	ELSIF TRUE 	
	AND fbPis.m_CheckByRecipe(stPis:=stPis_Tank_Water, 			req:=E_Piston_Recipe_State.Release)
	AND fbPis.m_CheckByRecipe(stPis:=stPis_Tank_R_Water, 		req:=E_Piston_Recipe_State.Release)
	AND fbPis.m_CheckByRecipe(stPis:=stPis_Tank_Detergent, 		req:=E_Piston_Recipe_State.Release)
	AND fbPis.m_CheckByRecipe(stPis:=stPis_Tank_DisInfection, 	req:=E_Piston_Recipe_State.Act)
	AND fbPis.m_CheckByRecipe(stPis:=stPis_Drain, 				req:=E_Piston_Recipe_State.Act)
	THEN;
		eStatus:=E_CIP_Source.eT91_Sanitation;
	ELSE;
		eStatus:=E_CIP_Source.eNone;
	END_IF
ELSE;
	eStatus:=E_CIP_Source.eNone;
END_IF
END_ACTION

METHOD m_CheckStatus : BOOL
VAR_INPUT
	eReqStatus		: E_CIP_Source;
END_VAR
IF eStatus=eReqStatus 
AND eProcess=E_CIP_Source.eNone
AND eReq=E_CIP_Source.eNone
AND bReady
AND bDone
AND NOT bRun
THEN;
	m_CheckStatus:=TRUE;
END_IF
END_METHOD

METHOD m_IsFree : BOOL
// In Ready with no request: a command given now will not be lost
IF eProcess=E_CIP_Source.eNone
AND eReq=E_CIP_Source.eNone
AND bReady
AND NOT bRun
THEN;
	m_IsFree:=TRUE;
END_IF
END_METHOD

METHOD m_Request_Reset : BOOL
VAR_IN_OUT
	memo: R_TRIG;
END_VAR
memo(CLK:=eReq=0);
IF TRUE 
AND memo.Q
THEN;
	SFCReset:=TRUE;
END_IF
END_METHOD

METHOD m_Run : BOOL
VAR_INPUT
	eReqProc			: E_CIP_Source;
END_VAR
IF eProcess=E_CIP_Source.eNone THEN;
	eProcess:=eReq:=eReqProc;
	bDone:=FALSE;
	m_Run:=TRUE;
END_IF
END_METHOD

METHOD m_Set_SFCFlags_Reference : BOOL
//Set reference to SFC flags

refSFC.SFCInit REF= SFCInit;
refSFC.SFCReset REF= SFCReset;
refSFC.SFCError REF= SFCError;
refSFC.SFCEnableLimit REF= SFCEnableLimit;
refSFC.SFCErrorStep REF= SFCErrorStep;
refSFC.SFCErrorPOU REF= SFCErrorPOU;
refSFC.SFCQuitError REF= SFCQuitError;
refSFC.SFCPause REF= SFCPause;
refSFC.SFCTrans REF= SFCTrans;
refSFC.SFCCurrentStep REF= SFCCurrentStep;
refSFC.SFCTip REF= SFCTip;
refSFC.SFCTipMode REF= SFCTipMode;

// Cycle handle for SFC
m_SFC_Handle();
END_METHOD

END_FUNCTION_BLOCK

// ---- 00 Library/03 SFC/FB_SFC_Cycle.TcPOU
FUNCTION_BLOCK FB_SFC_Cycle
VAR_INPUT

END_VAR
VAR_OUTPUT
END_VAR
VAR
	refSFC: ST_SFC;

	bInit: BOOL;
	bResetCycle: BOOL;
	bResume: BOOL;
	bRun: BOOL;	
	bReady: BOOL;
	bDone: BOOL;
	bToBe_Done: BOOL;
	
	bStepMode: BOOL;
	bNextStep: BOOL;



	bStepDone: BOOL;
	ton_StepTime: TON;
	
	StageDelayByRecipe: TIME;
	
	//fbPis_Meth: FB_Piston;

	rtDone	: R_TRIG;
	rtRun	: R_TRIG;
	sLastStepBefore_Error	: STRING;
	sError_Message			: STRING;
	
	ErrorSFC: BOOL;

	tonResetCycle: TON;
	
	stMode_zone	: REFERENCE TO ST_Mode;
	stOper_zone	: REFERENCE TO ST_OperationButtons;
	ftStateSafe : F_TRIG;
	
END_VAR

METHOD m_Reset_LastStepBeforeError : BOOL
VAR_INPUT
END_VAR
sLastStepBefore_Error:='';
END_METHOD

METHOD m_Set_LastStepBeforeError : BOOL
VAR_INPUT
END_VAR
sLastStepBefore_Error:=refSFC.SFCCurrentStep;
END_METHOD

METHOD m_Set_Mode_Reference : BOOL
VAR_INPUT
	inMoedeZone: E_ModeZone;
END_VAR
stMode_zone REF=(stMode[inMoedeZone]);
stOper_zone REF=(stOper[inMoedeZone]);
END_METHOD

METHOD m_SFC_Handle : BOOL
VAR_INPUT
END_VAR

VAR
	
END_VAR
IF NOT __ISVALIDREF(refSFC.SFCInit) 
OR NOT  __ISVALIDREF(refSFC.SFCReset) 
OR NOT  __ISVALIDREF(refSFC.SFCError) 
OR NOT  __ISVALIDREF(refSFC.SFCEnableLimit) 
OR NOT  __ISVALIDREF(refSFC.SFCErrorStep) 
OR NOT  __ISVALIDREF(refSFC.SFCErrorPOU) 
OR NOT  __ISVALIDREF(refSFC.SFCQuitError) 
OR NOT  __ISVALIDREF(refSFC.SFCPause) 
OR NOT  __ISVALIDREF(refSFC.SFCTrans) 
OR NOT  __ISVALIDREF(refSFC.SFCCurrentStep) 
OR NOT  __ISVALIDREF(refSFC.SFCTip) 
OR NOT  __ISVALIDREF(refSFC.SFCTipMode) 
THEN;
	RETURN;
END_IF

refSFC.SFCEnableLimit:=TRUE;
IF refSFC.SFCTrans THEN;
	bStepDone:=FALSE;
	ton_StepTime(IN:=FALSE);
ELSE;
	ton_StepTime(IN:=TRUE); //depend on step condition
END_IF

IF bInit THEN;
	refSFC.SFCInit:=TRUE;
ELSE;
	refSFC.SFCInit:=FALSE;
END_IF

IF refSFC.SFCError THEN;
	refSFC.SFCPause:=TRUE;
	ErrorSFC:=TRUE;
	m_Set_LastStepBeforeError();
END_IF

IF refSFC.SFCQuitError THEN;
	refSFC.SFCPause:=FALSE;
	ErrorSFC:=FALSE;
	refSFC.SFCQuitError:=FALSE;
	m_Reset_LastStepBeforeError();
	sError_Message:='';
END_IF

IF refSFC.SFCCurrentStep='Ready' THEN;
	bReady:=TRUE;
ELSE;
	bReady:=FALSE;
END_IF

rtDone(CLK:=refSFC.SFCCurrentStep='Done');
IF rtDone.Q THEN;
	bDone:=TRUE;
END_IF
rtRun(CLK:=bRun);
IF rtRun.Q THEN;
	bDone:=FALSE;
END_IF

IF bResume THEN;
	ErrorSFC:=FALSE;
	refSFC.SFCError:=FALSE;
	refSFC.SFCPause:=FALSE;
	m_Reset_LastStepBeforeError();
	bResume:=FALSE;
END_IF


tonResetCycle(PT:=T#0.5S,IN:=bResetCycle);
IF bResetCycle THEN;
	refSFC.SFCReset:=TRUE;
	//tonResetCycle.IN:=TRUE;
END_IF
IF tonResetCycle.Q THEN;
	bResetCycle:=FALSE;
	refSFC.SFCReset:=FALSE;
END_IF

StepByStep();

IF NOT __ISVALIDREF(stMode_zone)
OR NOT __ISVALIDREF(stOper_zone)
THEN;
	RETURN;
ELSE;
	//IF prg_Safety.ftStateSafe.Q THEN;
	ftStateSafe(CLK:=stMode_zone.bStateSafe_mode);
	IF ftStateSafe.Q THEN;
		//bResetCycle:=TRUE;
	END_IF	
END_IF



(*
rtDone(CLK:=bDone);
IF rtDone.Q THEN
	bToBe_Done:=FALSE;
END_IF
*)
END_METHOD

METHOD mInit : BOOL
VAR_INPUT
END_VAR
bInit:=TRUE;
bToBe_Done:=FALSE;
END_METHOD

METHOD mResetCycle : BOOL
VAR_INPUT
END_VAR
bResetCycle:=TRUE;
bRun:=FALSE;
refSFC.SFCReset:=TRUE;
END_METHOD

METHOD mRun : BOOL
VAR_INPUT
	
END_VAR
bRun:=TRUE;
bDone:=FALSE;

IF rtDone.Q THEN;
	mRun:=TRUE;	
END_IF
END_METHOD

METHOD mToBe_Done : BOOL
VAR_INPUT
END_VAR
bToBe_Done:=TRUE;
bDone:=FALSE;
END_METHOD

METHOD StepByStep : BOOL
VAR_INPUT
END_VAR


IF bStepMode THEN;
	IF refSFC.SFCTrans THEN;
		refSFC.SFCTipMode:=TRUE;
		bNextStep:=FALSE;
	END_IF
	IF bNextStep THEN;
		refSFC.SFCTipMode:=FALSE;
	END_IF
ELSE;
	refSFC.SFCTipMode:=FALSE;
END_IF
END_METHOD

END_FUNCTION_BLOCK

// ---- 03 Project/23 CIP/FB_CIP_Return.TcPOU
FUNCTION_BLOCK FB_CIP_Return EXTENDS FB_SFC_Cycle IMPLEMENTS ITF_FB_SFC_Cycle
VAR_INPUT
	//eElementID			: E_Element_List;
	
	valTank_Water			: E_Pis_Name;
	valTank_Water_1			: E_Pis_Name;
	valTank_R_Water			: E_Pis_Name;
	valTank_R_Water_1		: E_Pis_Name;
	valTank_Detergent		: E_Pis_Name;
	valTank_Detergent_1		: E_Pis_Name;
	valTank_DisInfection	: E_Pis_Name;
	valTank_DisInfection_1	: E_Pis_Name;
	valDrain				: E_Pis_Name;
	
END_VAR
VAR_OUTPUT
END_VAR
VAR
	//refElement		: REFERENCE TO FB_Element;
	//refState_Long		: REFERENCE TO E_Element_State_Long;
	eReq				: E_CIP_Return;
	eProcess			: E_CIP_Return;
	eStatus				: E_CIP_Return;
	
	fbPis						: FB_Piston;
	stPis_Tank_Water			: REFERENCE TO ST_Piston;
	stPis_Tank_Water_1			: REFERENCE TO ST_Piston;
	stPis_Tank_R_Water			: REFERENCE TO ST_Piston;
	stPis_Tank_R_Water_1		: REFERENCE TO ST_Piston;
	stPis_Tank_Detergent		: REFERENCE TO ST_Piston;
	stPis_Tank_Detergent_1		: REFERENCE TO ST_Piston;
	stPis_Tank_DisInfection		: REFERENCE TO ST_Piston;
	stPis_Tank_DisInfection_1	: REFERENCE TO ST_Piston;
	stPis_Drain					: REFERENCE TO ST_Piston;
	rt_Req_Reset: R_TRIG;
END_VAR
VAR_IN_OUT


END_VAR

act_GetReference();

act_Oper();
IF NOT Init.x THEN;
	act_Status();
END_IF

m_Request_Reset(memo:=rt_Req_Reset);//

ACTION _aDetergent_active:
bStepDone:=FALSE;
IF TRUE 
AND eStatus=E_CIP_Return.eT92_Detergent
THEN;
	bStepDone:=TRUE;
END_IF
END_ACTION

ACTION _aDetergent_entry:
fbPis.m_SetByRecipe(stPis:=stPis_Tank_Water, 			req:=E_Piston_Recipe_State.Release);
fbPis.m_SetByRecipe(stPis:=stPis_Tank_Water_1, 			req:=E_Piston_Recipe_State.Release);
fbPis.m_SetByRecipe(stPis:=stPis_Tank_R_Water, 			req:=E_Piston_Recipe_State.Release);
fbPis.m_SetByRecipe(stPis:=stPis_Tank_R_Water_1, 		req:=E_Piston_Recipe_State.Release);
fbPis.m_SetByRecipe(stPis:=stPis_Tank_Detergent, 		req:=E_Piston_Recipe_State.Act);
fbPis.m_SetByRecipe(stPis:=stPis_Tank_Detergent_1, 		req:=E_Piston_Recipe_State.Act);
fbPis.m_SetByRecipe(stPis:=stPis_Tank_DisInfection_1, 	req:=E_Piston_Recipe_State.Release);
fbPis.m_SetByRecipe(stPis:=stPis_Tank_DisInfection, 	req:=E_Piston_Recipe_State.Release);
fbPis.m_SetByRecipe(stPis:=stPis_Drain, 				req:=E_Piston_Recipe_State.Release);
END_ACTION

ACTION _aDone_entry:
eProcess:=E_CIP_Return.eNone; 
eReq:=E_CIP_Return.eNone;
bRun:=FALSE;
bDone:=TRUE;
END_ACTION

ACTION _aDrain_active:
bStepDone:=FALSE;
IF TRUE 
AND eStatus=E_CIP_Return.eDrain
THEN;
	bStepDone:=TRUE;
END_IF
END_ACTION

ACTION _aDrain_entry:
fbPis.m_SetByRecipe(stPis:=stPis_Tank_Water, 			req:=E_Piston_Recipe_State.Release);
fbPis.m_SetByRecipe(stPis:=stPis_Tank_Water_1, 			req:=E_Piston_Recipe_State.Release);
fbPis.m_SetByRecipe(stPis:=stPis_Tank_R_Water, 			req:=E_Piston_Recipe_State.Release);
fbPis.m_SetByRecipe(stPis:=stPis_Tank_R_Water_1, 		req:=E_Piston_Recipe_State.Release);
fbPis.m_SetByRecipe(stPis:=stPis_Tank_Detergent, 		req:=E_Piston_Recipe_State.Release);
fbPis.m_SetByRecipe(stPis:=stPis_Tank_Detergent_1, 		req:=E_Piston_Recipe_State.Release);
fbPis.m_SetByRecipe(stPis:=stPis_Tank_DisInfection, 	req:=E_Piston_Recipe_State.Release);
fbPis.m_SetByRecipe(stPis:=stPis_Tank_DisInfection_1, 	req:=E_Piston_Recipe_State.Release);
fbPis.m_SetByRecipe(stPis:=stPis_Drain, 				req:=E_Piston_Recipe_State.Release);
END_ACTION

ACTION _aInit_active:
SFCReset:=FALSE;
END_ACTION

ACTION _aInit_exit:
eProcess:=E_CIP_Return.eNone;
eReq:=E_CIP_Return.eNone;
END_ACTION

ACTION _aR_Water_active:
bStepDone:=FALSE;
IF TRUE 
AND eStatus=E_CIP_Return.eT93_R_Water
THEN;
	bStepDone:=TRUE;
END_IF
END_ACTION

ACTION _aR_Water_entry:
fbPis.m_SetByRecipe(stPis:=stPis_Tank_Water, 			req:=E_Piston_Recipe_State.Release);
fbPis.m_SetByRecipe(stPis:=stPis_Tank_Water_1, 			req:=E_Piston_Recipe_State.Release);
fbPis.m_SetByRecipe(stPis:=stPis_Tank_R_Water, 			req:=E_Piston_Recipe_State.Act);
fbPis.m_SetByRecipe(stPis:=stPis_Tank_R_Water_1, 		req:=E_Piston_Recipe_State.Act);
fbPis.m_SetByRecipe(stPis:=stPis_Tank_Detergent, 		req:=E_Piston_Recipe_State.Release);
fbPis.m_SetByRecipe(stPis:=stPis_Tank_Detergent_1, 		req:=E_Piston_Recipe_State.Release);
fbPis.m_SetByRecipe(stPis:=stPis_Tank_DisInfection, 	req:=E_Piston_Recipe_State.Release);
fbPis.m_SetByRecipe(stPis:=stPis_Tank_DisInfection_1, 	req:=E_Piston_Recipe_State.Release);
fbPis.m_SetByRecipe(stPis:=stPis_Drain, 				req:=E_Piston_Recipe_State.Release);
END_ACTION

ACTION _aReady_active:


CASE eReq OF
	E_CIP_Return.eDrain:;
			IF TRUE THEN;
				eProcess:=E_CIP_Return.eDrain;
			END_IF

	E_CIP_Return.eT91_Sanitation:;
			IF TRUE THEN;
				eProcess:=E_CIP_Return.eT91_Sanitation;
			END_IF	
			
	E_CIP_Return.eT92_Detergent:;
			IF TRUE THEN;
				eProcess:=E_CIP_Return.eT92_Detergent;
			END_IF	

	E_CIP_Return.eT93_R_Water:;
			IF TRUE THEN;
				eProcess:=E_CIP_Return.eT93_R_Water;
			END_IF	
			
	E_CIP_Return.eT94_Water:;
			IF TRUE THEN;
				eProcess:=E_CIP_Return.eT94_Water;
			END_IF	

END_CASE
END_ACTION

ACTION _aReady_entry:

END_ACTION

ACTION _aReady_exit:
bRun:=TRUE;
bDone:=FALSE;
END_ACTION

ACTION _aSanitation_active:
bStepDone:=FALSE;
IF TRUE 
AND eStatus=E_CIP_Return.eT91_Sanitation
THEN;
	bStepDone:=TRUE;
END_IF
END_ACTION

ACTION _aSanitation_entry:
fbPis.m_SetByRecipe(stPis:=stPis_Tank_Water, 			req:=E_Piston_Recipe_State.Release);
fbPis.m_SetByRecipe(stPis:=stPis_Tank_Water_1, 			req:=E_Piston_Recipe_State.Release);
fbPis.m_SetByRecipe(stPis:=stPis_Tank_R_Water, 			req:=E_Piston_Recipe_State.Release);
fbPis.m_SetByRecipe(stPis:=stPis_Tank_R_Water_1, 		req:=E_Piston_Recipe_State.Release);
fbPis.m_SetByRecipe(stPis:=stPis_Tank_Detergent, 		req:=E_Piston_Recipe_State.Release);
fbPis.m_SetByRecipe(stPis:=stPis_Tank_Detergent_1, 		req:=E_Piston_Recipe_State.Release);
fbPis.m_SetByRecipe(stPis:=stPis_Tank_DisInfection, 	req:=E_Piston_Recipe_State.Act);
fbPis.m_SetByRecipe(stPis:=stPis_Tank_DisInfection_1, 	req:=E_Piston_Recipe_State.Act);
fbPis.m_SetByRecipe(stPis:=stPis_Drain, 				req:=E_Piston_Recipe_State.Release);
END_ACTION

ACTION _aWater_active:
bStepDone:=FALSE;
IF TRUE 
AND eStatus=E_CIP_Return.eT94_Water
THEN;
	bStepDone:=TRUE;
END_IF
END_ACTION

ACTION _aWater_entry:
fbPis.m_SetByRecipe(stPis:=stPis_Tank_Water, 			req:=E_Piston_Recipe_State.Act);
fbPis.m_SetByRecipe(stPis:=stPis_Tank_Water_1, 			req:=E_Piston_Recipe_State.Act);
fbPis.m_SetByRecipe(stPis:=stPis_Tank_R_Water, 			req:=E_Piston_Recipe_State.Release);
fbPis.m_SetByRecipe(stPis:=stPis_Tank_R_Water_1, 		req:=E_Piston_Recipe_State.Release);
fbPis.m_SetByRecipe(stPis:=stPis_Tank_Detergent, 		req:=E_Piston_Recipe_State.Release);
fbPis.m_SetByRecipe(stPis:=stPis_Tank_Detergent_1, 		req:=E_Piston_Recipe_State.Release);
fbPis.m_SetByRecipe(stPis:=stPis_Tank_DisInfection, 	req:=E_Piston_Recipe_State.Release);
fbPis.m_SetByRecipe(stPis:=stPis_Tank_DisInfection_1, 	req:=E_Piston_Recipe_State.Release);
fbPis.m_SetByRecipe(stPis:=stPis_Drain, 				req:=E_Piston_Recipe_State.Act);
END_ACTION

ACTION act_GetReference:
m_Set_SFCFlags_Reference();
//refElement REF= fbElement[eElementID];
//refState_Long REF= fbElement[eElementID].eState_Long;
	
stPis_Tank_Water				REF= g_Piston.stPis[valTank_Water];
stPis_Tank_Water_1				REF= g_Piston.stPis[valTank_Water_1];
stPis_Tank_R_Water				REF= g_Piston.stPis[valTank_R_Water];
stPis_Tank_R_Water_1			REF= g_Piston.stPis[valTank_R_Water_1];
stPis_Tank_Detergent			REF= g_Piston.stPis[valTank_Detergent];
stPis_Tank_Detergent_1			REF= g_Piston.stPis[valTank_Detergent_1];
stPis_Tank_DisInfection			REF= g_Piston.stPis[valTank_DisInfection];
stPis_Tank_DisInfection_1		REF= g_Piston.stPis[valTank_DisInfection_1];
stPis_Drain						REF= g_Piston.stPis[valDrain];
END_ACTION

ACTION act_Oper:
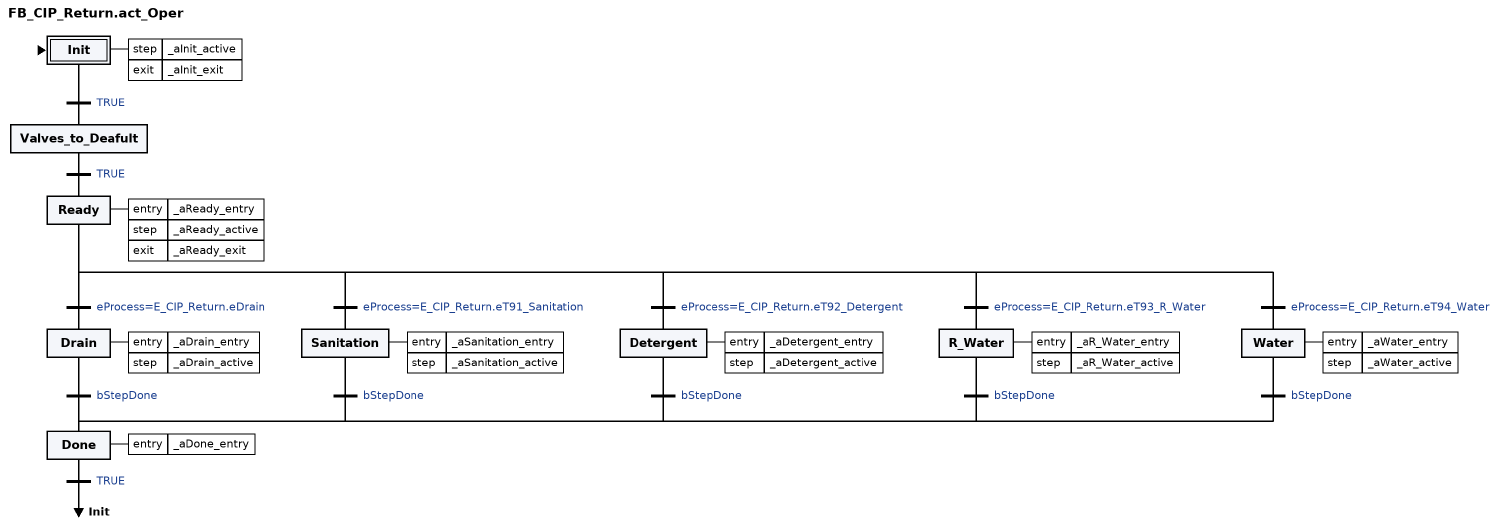
INITIAL_STEP Init:  // min time T#0.5s
    _aInit_active(N);  // step action
    _aInit_exit(P0);  // exit action
END_STEP
TRANSITION FROM Init TO Valves_to_Deafult
    := TRUE;
END_TRANSITION
STEP Valves_to_Deafult:
END_STEP
TRANSITION FROM Valves_to_Deafult TO Ready
    := TRUE;
END_TRANSITION
STEP Ready:
    _aReady_entry(P1);  // entry action
    _aReady_active(N);  // step action
    _aReady_exit(P0);  // exit action
END_STEP
TRANSITION FROM Ready TO Drain
    := eProcess=E_CIP_Return.eDrain;
END_TRANSITION
STEP Drain:
    _aDrain_entry(P1);  // entry action
    _aDrain_active(N);  // step action
END_STEP
TRANSITION FROM Drain TO Done
    := bStepDone;
END_TRANSITION
TRANSITION FROM Ready TO Sanitation
    := eProcess=E_CIP_Return.eT91_Sanitation;
END_TRANSITION
STEP Sanitation:
    _aSanitation_entry(P1);  // entry action
    _aSanitation_active(N);  // step action
END_STEP
TRANSITION FROM Sanitation TO Done
    := bStepDone;
END_TRANSITION
TRANSITION FROM Ready TO Detergent
    := eProcess=E_CIP_Return.eT92_Detergent;
END_TRANSITION
STEP Detergent:
    _aDetergent_entry(P1);  // entry action
    _aDetergent_active(N);  // step action
END_STEP
TRANSITION FROM Detergent TO Done
    := bStepDone;
END_TRANSITION
TRANSITION FROM Ready TO R_Water
    := eProcess=E_CIP_Return.eT93_R_Water;
END_TRANSITION
STEP R_Water:
    _aR_Water_entry(P1);  // entry action
    _aR_Water_active(N);  // step action
END_STEP
TRANSITION FROM R_Water TO Done
    := bStepDone;
END_TRANSITION
TRANSITION FROM Ready TO Water
    := eProcess=E_CIP_Return.eT94_Water;
END_TRANSITION
STEP Water:
    _aWater_entry(P1);  // entry action
    _aWater_active(N);  // step action
END_STEP
TRANSITION FROM Water TO Done
    := bStepDone;
END_TRANSITION
STEP Done:  // min time T#0.2s
    _aDone_entry(P1);  // entry action
END_STEP
TRANSITION FROM Done TO Init
    := TRUE;
END_TRANSITION
// branch label Branch1_act_Oper
END_ACTION

ACTION act_Status:
IF bReady AND bDone OR TRUE THEN;
	IF TRUE 
	AND fbPis.m_CheckByRecipe(stPis:=stPis_Tank_Water, 			req:=E_Piston_Recipe_State.Release)
	AND fbPis.m_CheckByRecipe(stPis:=stPis_Tank_R_Water, 		req:=E_Piston_Recipe_State.Release)
	AND fbPis.m_CheckByRecipe(stPis:=stPis_Tank_Detergent, 		req:=E_Piston_Recipe_State.Release)
	AND fbPis.m_CheckByRecipe(stPis:=stPis_Tank_DisInfection, 	req:=E_Piston_Recipe_State.Release)
	AND fbPis.m_CheckByRecipe(stPis:=stPis_Drain, 				req:=E_Piston_Recipe_State.Release)
	AND fbPis.m_CheckByRecipe(stPis:=stPis_Tank_Water_1, 		req:=E_Piston_Recipe_State.Release)
	AND fbPis.m_CheckByRecipe(stPis:=stPis_Tank_R_Water_1, 		req:=E_Piston_Recipe_State.Release)
	AND fbPis.m_CheckByRecipe(stPis:=stPis_Tank_Detergent_1, 	req:=E_Piston_Recipe_State.Release)
	AND fbPis.m_CheckByRecipe(stPis:=stPis_Tank_DisInfection_1, req:=E_Piston_Recipe_State.Release)
	THEN;
		eStatus:=E_CIP_Return.eDrain;
	
	ELSIF TRUE 
	AND fbPis.m_CheckByRecipe(stPis:=stPis_Tank_Water, 			req:=E_Piston_Recipe_State.Act)
	AND fbPis.m_CheckByRecipe(stPis:=stPis_Tank_R_Water, 		req:=E_Piston_Recipe_State.Release)
	AND fbPis.m_CheckByRecipe(stPis:=stPis_Tank_Detergent, 		req:=E_Piston_Recipe_State.Release)
	AND fbPis.m_CheckByRecipe(stPis:=stPis_Tank_DisInfection, 	req:=E_Piston_Recipe_State.Release)
	AND fbPis.m_CheckByRecipe(stPis:=stPis_Drain, 				req:=E_Piston_Recipe_State.Act)
	AND fbPis.m_CheckByRecipe(stPis:=stPis_Tank_Water_1, 		req:=E_Piston_Recipe_State.Act)
	AND fbPis.m_CheckByRecipe(stPis:=stPis_Tank_R_Water_1, 		req:=E_Piston_Recipe_State.Release)
	AND fbPis.m_CheckByRecipe(stPis:=stPis_Tank_Detergent_1, 	req:=E_Piston_Recipe_State.Release)
	AND fbPis.m_CheckByRecipe(stPis:=stPis_Tank_DisInfection_1, req:=E_Piston_Recipe_State.Release)
	THEN;
		eStatus:=E_CIP_Return.eT94_Water;
		
	ELSIF TRUE 
	AND fbPis.m_CheckByRecipe(stPis:=stPis_Tank_Water, 			req:=E_Piston_Recipe_State.Release)
	AND fbPis.m_CheckByRecipe(stPis:=stPis_Tank_R_Water, 		req:=E_Piston_Recipe_State.Act)
	AND fbPis.m_CheckByRecipe(stPis:=stPis_Tank_Detergent, 		req:=E_Piston_Recipe_State.Release)
	AND fbPis.m_CheckByRecipe(stPis:=stPis_Tank_DisInfection, 	req:=E_Piston_Recipe_State.Release)
	AND fbPis.m_CheckByRecipe(stPis:=stPis_Drain, 				req:=E_Piston_Recipe_State.Release)
	AND fbPis.m_CheckByRecipe(stPis:=stPis_Tank_Water_1, 			req:=E_Piston_Recipe_State.Release)
	AND fbPis.m_CheckByRecipe(stPis:=stPis_Tank_R_Water_1, 			req:=E_Piston_Recipe_State.Act)
	AND fbPis.m_CheckByRecipe(stPis:=stPis_Tank_Detergent_1, 		req:=E_Piston_Recipe_State.Release)
	AND fbPis.m_CheckByRecipe(stPis:=stPis_Tank_DisInfection_1, 	req:=E_Piston_Recipe_State.Release)
	THEN;
		eStatus:=E_CIP_Return.eT93_R_Water;
		
	ELSIF TRUE 	
	AND fbPis.m_CheckByRecipe(stPis:=stPis_Tank_Water, 			req:=E_Piston_Recipe_State.Release)
	AND fbPis.m_CheckByRecipe(stPis:=stPis_Tank_R_Water, 		req:=E_Piston_Recipe_State.Release)
	AND fbPis.m_CheckByRecipe(stPis:=stPis_Tank_Detergent, 		req:=E_Piston_Recipe_State.Act)
	AND fbPis.m_CheckByRecipe(stPis:=stPis_Tank_DisInfection, 	req:=E_Piston_Recipe_State.Release)
	AND fbPis.m_CheckByRecipe(stPis:=stPis_Drain, 				req:=E_Piston_Recipe_State.Release)
	AND fbPis.m_CheckByRecipe(stPis:=stPis_Tank_Water_1, 			req:=E_Piston_Recipe_State.Release)
	AND fbPis.m_CheckByRecipe(stPis:=stPis_Tank_R_Water_1, 			req:=E_Piston_Recipe_State.Release)
	AND fbPis.m_CheckByRecipe(stPis:=stPis_Tank_Detergent_1, 		req:=E_Piston_Recipe_State.Act)
	AND fbPis.m_CheckByRecipe(stPis:=stPis_Tank_DisInfection_1, 	req:=E_Piston_Recipe_State.Release)
	THEN;
		eStatus:=E_CIP_Return.eT92_Detergent;
		
	ELSIF TRUE 	
	AND fbPis.m_CheckByRecipe(stPis:=stPis_Tank_Water, 			req:=E_Piston_Recipe_State.Release)
	AND fbPis.m_CheckByRecipe(stPis:=stPis_Tank_R_Water, 		req:=E_Piston_Recipe_State.Release)
	AND fbPis.m_CheckByRecipe(stPis:=stPis_Tank_Detergent, 		req:=E_Piston_Recipe_State.Release)
	AND fbPis.m_CheckByRecipe(stPis:=stPis_Tank_DisInfection, 	req:=E_Piston_Recipe_State.Act)
	AND fbPis.m_CheckByRecipe(stPis:=stPis_Drain, 				req:=E_Piston_Recipe_State.Release)
	AND fbPis.m_CheckByRecipe(stPis:=stPis_Tank_Water_1, 			req:=E_Piston_Recipe_State.Release)
	AND fbPis.m_CheckByRecipe(stPis:=stPis_Tank_R_Water_1, 			req:=E_Piston_Recipe_State.Release)
	AND fbPis.m_CheckByRecipe(stPis:=stPis_Tank_Detergent_1, 		req:=E_Piston_Recipe_State.Release)
	AND fbPis.m_CheckByRecipe(stPis:=stPis_Tank_DisInfection_1, 	req:=E_Piston_Recipe_State.Act)
	THEN;
		eStatus:=E_CIP_Return.eT91_Sanitation;
	ELSE;
		eStatus:=E_CIP_Return.eNone;
	END_IF
ELSE;
	eStatus:=E_CIP_Return.eNone;
END_IF
END_ACTION

METHOD m_CheckStatus : BOOL
VAR_INPUT
	eReqStatus		: E_CIP_Return;
END_VAR
IF eStatus=eReqStatus 
AND eProcess=E_CIP_Return.eNone
AND eReq=E_CIP_Return.eNone
AND bReady
AND bDone
AND NOT bRun
THEN;
	m_CheckStatus:=TRUE;
END_IF
END_METHOD

METHOD m_IsFree : BOOL
// In Ready with no request: a command given now will not be lost
IF eProcess=E_CIP_Return.eNone
AND eReq=E_CIP_Return.eNone
AND bReady
AND NOT bRun
THEN;
	m_IsFree:=TRUE;
END_IF
END_METHOD

METHOD m_Request_Reset : BOOL
VAR_IN_OUT
	memo: R_TRIG;
END_VAR
memo(CLK:=eReq=0);
IF TRUE 
AND memo.Q
THEN;
	SFCReset:=TRUE;
END_IF
END_METHOD

METHOD m_Run : BOOL
VAR_INPUT
	eReqProc			: E_CIP_Return;
END_VAR
IF eProcess=E_CIP_Return.eNone THEN;
	eProcess:=eReq:=eReqProc;
	bDone:=FALSE;
	m_Run:=TRUE;
END_IF
END_METHOD

METHOD m_Set_SFCFlags_Reference : BOOL
//Set reference to SFC flags

refSFC.SFCInit REF= SFCInit;
refSFC.SFCReset REF= SFCReset;
refSFC.SFCError REF= SFCError;
refSFC.SFCEnableLimit REF= SFCEnableLimit;
refSFC.SFCErrorStep REF= SFCErrorStep;
refSFC.SFCErrorPOU REF= SFCErrorPOU;
refSFC.SFCQuitError REF= SFCQuitError;
refSFC.SFCPause REF= SFCPause;
refSFC.SFCTrans REF= SFCTrans;
refSFC.SFCCurrentStep REF= SFCCurrentStep;
refSFC.SFCTip REF= SFCTip;
refSFC.SFCTipMode REF= SFCTipMode;

// Cycle handle for SFC
m_SFC_Handle();
END_METHOD

END_FUNCTION_BLOCK

// ---- 03 Project/23 CIP/FB_CIP_Client.TcPOU
FUNCTION_BLOCK FB_CIP_Client EXTENDS FB_SFC_Cycle IMPLEMENTS ITF_FB_SFC_Cycle
VAR_INPUT
	//eElementID			: E_Element_List;
	
	valClient_Source		: E_Pis_Name;
	valClient_Return		: E_Pis_Name;
	valS_Marinade_Up		: E_Pis_Name;
	//valS_Marinade_Up_Drain	: E_Pis_Name;
	valS_Marinade_Low		: E_Pis_Name;
	valS_Color_Up			: E_Pis_Name;
	//valS_Color_Up_Drain		: E_Pis_Name;
	valS_Color_Low			: E_Pis_Name;
	//valTank_1				: E_Pis_Name;
	//valTank_2				: E_Pis_Name;
	//valTank_3				: E_Pis_Name;
	//valTank_4				: E_Pis_Name;
	//valS_Marinade_Low_Select	: E_Pis_Name;
	//valS_Color_Low_Select	: E_Pis_Name;
	valDrain				: E_Pis_Name;
	valLoop					: E_Pis_Name;//V1030
	valS_Future				: E_Pis_Name;
	
END_VAR
VAR_OUTPUT
END_VAR
VAR
	//refElement		: REFERENCE TO FB_Element;
	//refState_Long		: REFERENCE TO E_Element_State_Long;
	eReq				: E_CIP_Client_Selector;
	eProcess			: E_CIP_Client_Selector;
	eStatus				: E_CIP_Client_Selector;
	
	fbPis					: FB_Piston;
	stPis_Client_Source			: REFERENCE TO ST_Piston;
	stPis_Client_Return			: REFERENCE TO ST_Piston;
	stPis_S_Marinade_Up			: REFERENCE TO ST_Piston;
	//stPis_S_Marinade_Up_Drain	: REFERENCE TO ST_Piston;
	stPis_S_Marinade_Low		: REFERENCE TO ST_Piston;
	stPis_S_Color_Up			: REFERENCE TO ST_Piston;
	//stPis_S_Color_Up_Drain		: REFERENCE TO ST_Piston;
	stPis_S_Color_Low			: REFERENCE TO ST_Piston;
	//stPis_Tank_1				: REFERENCE TO ST_Piston;
	//stPis_Tank_2				: REFERENCE TO ST_Piston;
	//stPis_Tank_3				: REFERENCE TO ST_Piston;
	//stPis_Tank_4				: REFERENCE TO ST_Piston;
	//stPis_S_Marinade_Low_Select	: REFERENCE TO ST_Piston;
	//stPis_S_Color_Low_Select	: REFERENCE TO ST_Piston;
	stPis_Drain					: REFERENCE TO ST_Piston;	
	stPis_Loop					: REFERENCE TO ST_Piston;//V1030
	stPis_S_Future				: REFERENCE TO ST_Piston;

	tonDrainTime: TON;
	
	rt_Req_Reset: R_TRIG;

END_VAR
VAR_IN_OUT


END_VAR

act_GetReference();

act_Oper();
IF NOT Init.x THEN;
	act_Status();
END_IF

tonDrainTime(PT:=T#1M, IN:=eStatus=E_CIP_Client_Selector.eDrain);
IF tonDrainTime.Q 
AND eReq=E_CIP_Client_Selector.eNone
AND eProcess=E_CIP_Client_Selector.eNone
THEN;
	eReq:=E_CIP_Client_Selector.eClose;
END_IF

m_Request_Reset(memo:=rt_Req_Reset);//rt_Req_Reset: R_TRIG;

ACTION _aClose_active:
bStepDone:=FALSE;
IF TRUE 
AND eStatus=E_CIP_Client_Selector.eClose
THEN;
	bStepDone:=TRUE;
END_IF
END_ACTION

ACTION _aClose_entry:
fbPis.m_SetByRecipe(stPis:=stPis_Client_Source, 		req:=E_Piston_Recipe_State.Release);
fbPis.m_SetByRecipe(stPis:=stPis_Client_Return, 		req:=E_Piston_Recipe_State.Release);
fbPis.m_SetByRecipe(stPis:=stPis_S_Marinade_Up, 		req:=E_Piston_Recipe_State.Release);
fbPis.m_SetByRecipe(stPis:=stPis_S_Marinade_Low, 		req:=E_Piston_Recipe_State.Release);
fbPis.m_SetByRecipe(stPis:=stPis_S_Color_Up, 			req:=E_Piston_Recipe_State.Release);
fbPis.m_SetByRecipe(stPis:=stPis_S_Color_Low, 			req:=E_Piston_Recipe_State.Release);
fbPis.m_SetByRecipe(stPis:=stPis_Drain, 				req:=E_Piston_Recipe_State.Release);
fbPis.m_SetByRecipe(stPis:=stPis_Loop, 					req:=E_Piston_Recipe_State.Release);
fbPis.m_SetByRecipe(stPis:=stPis_S_Future, 				req:=E_Piston_Recipe_State.Release);
END_ACTION

ACTION _aColor_Low_active:
bStepDone:=FALSE;
IF TRUE 
AND eStatus=E_CIP_Client_Selector.eColor_Low
THEN;
	bStepDone:=TRUE;
END_IF
END_ACTION

ACTION _aColor_Low_entry:
fbPis.m_SetByRecipe(stPis:=stPis_Client_Source, 		req:=E_Piston_Recipe_State.Act);
fbPis.m_SetByRecipe(stPis:=stPis_Client_Return, 		req:=E_Piston_Recipe_State.Act);
fbPis.m_SetByRecipe(stPis:=stPis_S_Marinade_Up, 		req:=E_Piston_Recipe_State.Release);
fbPis.m_SetByRecipe(stPis:=stPis_S_Marinade_Low, 		req:=E_Piston_Recipe_State.Release);
fbPis.m_SetByRecipe(stPis:=stPis_S_Color_Up, 			req:=E_Piston_Recipe_State.Release);
fbPis.m_SetByRecipe(stPis:=stPis_S_Color_Low, 			req:=E_Piston_Recipe_State.Act);
fbPis.m_SetByRecipe(stPis:=stPis_Drain, 				req:=E_Piston_Recipe_State.Release);
fbPis.m_SetByRecipe(stPis:=stPis_Loop, 					req:=E_Piston_Recipe_State.Release);
fbPis.m_SetByRecipe(stPis:=stPis_S_Future, 				req:=E_Piston_Recipe_State.Release);
END_ACTION

ACTION _aColor_Up_active:
bStepDone:=FALSE;
IF TRUE 
AND eStatus=E_CIP_Client_Selector.eColor_Up
THEN;
	bStepDone:=TRUE;
END_IF
END_ACTION

ACTION _aColor_Up_entry:
fbPis.m_SetByRecipe(stPis:=stPis_Client_Source, 		req:=E_Piston_Recipe_State.Act);
fbPis.m_SetByRecipe(stPis:=stPis_Client_Return, 		req:=E_Piston_Recipe_State.Act);
fbPis.m_SetByRecipe(stPis:=stPis_S_Marinade_Up, 		req:=E_Piston_Recipe_State.Release);
fbPis.m_SetByRecipe(stPis:=stPis_S_Marinade_Low, 		req:=E_Piston_Recipe_State.Release);
fbPis.m_SetByRecipe(stPis:=stPis_S_Color_Up, 			req:=E_Piston_Recipe_State.Act);
fbPis.m_SetByRecipe(stPis:=stPis_S_Color_Low, 			req:=E_Piston_Recipe_State.Release);
fbPis.m_SetByRecipe(stPis:=stPis_Drain, 				req:=E_Piston_Recipe_State.Release);
fbPis.m_SetByRecipe(stPis:=stPis_Loop, 					req:=E_Piston_Recipe_State.Release);
fbPis.m_SetByRecipe(stPis:=stPis_S_Future, 				req:=E_Piston_Recipe_State.Release);
END_ACTION

ACTION _aDone_entry:
eProcess:=E_CIP_Usage.eNotInUse;
eReq:=E_CIP_Usage.eNotInUse;
bRun:=FALSE;
bDone:=TRUE;
END_ACTION

ACTION _aDrain_active:
bStepDone:=FALSE;
IF TRUE 
AND eStatus=E_CIP_Client_Selector.eDrain
THEN;
	bStepDone:=TRUE;
END_IF
END_ACTION

ACTION _aDrain_entry:
fbPis.m_SetByRecipe(stPis:=stPis_Client_Source, 		req:=E_Piston_Recipe_State.Release);
fbPis.m_SetByRecipe(stPis:=stPis_Client_Return, 		req:=E_Piston_Recipe_State.Release);
fbPis.m_SetByRecipe(stPis:=stPis_S_Marinade_Up, 		req:=E_Piston_Recipe_State.Release);
fbPis.m_SetByRecipe(stPis:=stPis_S_Marinade_Low, 		req:=E_Piston_Recipe_State.Release);
fbPis.m_SetByRecipe(stPis:=stPis_S_Color_Up, 			req:=E_Piston_Recipe_State.Release);
fbPis.m_SetByRecipe(stPis:=stPis_S_Color_Low, 			req:=E_Piston_Recipe_State.Release);
fbPis.m_SetByRecipe(stPis:=stPis_Drain, 				req:=E_Piston_Recipe_State.Act);
fbPis.m_SetByRecipe(stPis:=stPis_Loop, 					req:=E_Piston_Recipe_State.Release);
fbPis.m_SetByRecipe(stPis:=stPis_S_Future, 				req:=E_Piston_Recipe_State.Release);
END_ACTION

ACTION _aFuture_active:
bStepDone:=FALSE;
IF TRUE 
AND eStatus=E_CIP_Client_Selector.eFuture
THEN;
	bStepDone:=TRUE;
END_IF
END_ACTION

ACTION _aFuture_entry:
fbPis.m_SetByRecipe(stPis:=stPis_Client_Source, 		req:=E_Piston_Recipe_State.Act);
fbPis.m_SetByRecipe(stPis:=stPis_Client_Return, 		req:=E_Piston_Recipe_State.Act);
fbPis.m_SetByRecipe(stPis:=stPis_S_Marinade_Up, 		req:=E_Piston_Recipe_State.Release);
fbPis.m_SetByRecipe(stPis:=stPis_S_Marinade_Low, 		req:=E_Piston_Recipe_State.Release);
fbPis.m_SetByRecipe(stPis:=stPis_S_Color_Up, 			req:=E_Piston_Recipe_State.Release);
fbPis.m_SetByRecipe(stPis:=stPis_S_Color_Low, 			req:=E_Piston_Recipe_State.Release);
fbPis.m_SetByRecipe(stPis:=stPis_Drain, 				req:=E_Piston_Recipe_State.Release);
fbPis.m_SetByRecipe(stPis:=stPis_Loop, 					req:=E_Piston_Recipe_State.Release);
fbPis.m_SetByRecipe(stPis:=stPis_S_Future, 				req:=E_Piston_Recipe_State.Release);	//route to the plant: only source and return open
END_ACTION

ACTION _aInit_active:
SFCReset:=FALSE;
END_ACTION

ACTION _aInit_exit:
eProcess:=E_CIP_Usage.eNotInUse;
eReq:=E_CIP_Usage.eNotInUse;
END_ACTION

ACTION _aLoop_active:
bStepDone:=FALSE;
IF TRUE 
AND eStatus=E_CIP_Client_Selector.eLoop
THEN;
	bStepDone:=TRUE;
END_IF
END_ACTION

ACTION _aLoop_entry:
fbPis.m_SetByRecipe(stPis:=stPis_Client_Source, 		req:=E_Piston_Recipe_State.Act);
fbPis.m_SetByRecipe(stPis:=stPis_Client_Return, 		req:=E_Piston_Recipe_State.Act);
fbPis.m_SetByRecipe(stPis:=stPis_S_Marinade_Up, 		req:=E_Piston_Recipe_State.Release);
fbPis.m_SetByRecipe(stPis:=stPis_S_Marinade_Low, 		req:=E_Piston_Recipe_State.Release);
fbPis.m_SetByRecipe(stPis:=stPis_S_Color_Up, 			req:=E_Piston_Recipe_State.Release);
fbPis.m_SetByRecipe(stPis:=stPis_S_Color_Low, 			req:=E_Piston_Recipe_State.Release);
fbPis.m_SetByRecipe(stPis:=stPis_Drain, 				req:=E_Piston_Recipe_State.Act);
fbPis.m_SetByRecipe(stPis:=stPis_Loop, 					req:=E_Piston_Recipe_State.Act);
fbPis.m_SetByRecipe(stPis:=stPis_S_Future, 				req:=E_Piston_Recipe_State.Release);
END_ACTION

ACTION _aMarinade_Low_active:
bStepDone:=FALSE;
IF TRUE 
AND eStatus=E_CIP_Client_Selector.eMarinade_Low
THEN;
	bStepDone:=TRUE;
END_IF
END_ACTION

ACTION _aMarinade_Low_entry:
fbPis.m_SetByRecipe(stPis:=stPis_Client_Source, 		req:=E_Piston_Recipe_State.Act);
fbPis.m_SetByRecipe(stPis:=stPis_Client_Return, 		req:=E_Piston_Recipe_State.Act);
fbPis.m_SetByRecipe(stPis:=stPis_S_Marinade_Up, 		req:=E_Piston_Recipe_State.Release);
fbPis.m_SetByRecipe(stPis:=stPis_S_Marinade_Low, 		req:=E_Piston_Recipe_State.Act);
fbPis.m_SetByRecipe(stPis:=stPis_S_Color_Up, 			req:=E_Piston_Recipe_State.Release);
fbPis.m_SetByRecipe(stPis:=stPis_S_Color_Low, 			req:=E_Piston_Recipe_State.Release);
fbPis.m_SetByRecipe(stPis:=stPis_Drain, 				req:=E_Piston_Recipe_State.Release);
fbPis.m_SetByRecipe(stPis:=stPis_Loop, 					req:=E_Piston_Recipe_State.Release);
fbPis.m_SetByRecipe(stPis:=stPis_S_Future, 				req:=E_Piston_Recipe_State.Release);
END_ACTION

ACTION _aMarinade_Up_active:
bStepDone:=FALSE;
IF TRUE 
AND eStatus=E_CIP_Client_Selector.eMarinade_Up
THEN;
	bStepDone:=TRUE;
END_IF
END_ACTION

ACTION _aMarinade_Up_entry:
fbPis.m_SetByRecipe(stPis:=stPis_Client_Source, 		req:=E_Piston_Recipe_State.Act);
fbPis.m_SetByRecipe(stPis:=stPis_Client_Return, 		req:=E_Piston_Recipe_State.Act);
fbPis.m_SetByRecipe(stPis:=stPis_S_Marinade_Up, 		req:=E_Piston_Recipe_State.Act);
fbPis.m_SetByRecipe(stPis:=stPis_S_Marinade_Low, 		req:=E_Piston_Recipe_State.Release);
fbPis.m_SetByRecipe(stPis:=stPis_S_Color_Up, 			req:=E_Piston_Recipe_State.Release);
fbPis.m_SetByRecipe(stPis:=stPis_S_Color_Low, 			req:=E_Piston_Recipe_State.Release);
fbPis.m_SetByRecipe(stPis:=stPis_Drain, 				req:=E_Piston_Recipe_State.Release);
fbPis.m_SetByRecipe(stPis:=stPis_Loop, 					req:=E_Piston_Recipe_State.Release);
fbPis.m_SetByRecipe(stPis:=stPis_S_Future, 				req:=E_Piston_Recipe_State.Release);
END_ACTION

ACTION _aReady_active:


IF eReq<>E_CIP_Client_Selector.eNone THEN;
	IF eProcess=E_CIP_Client_Selector.eNone 
	THEN;
		eProcess:=eReq;
	ELSE;
		eReq:=E_CIP_Client_Selector.eNone;
	END_IF
END_IF

(*
CASE eReq OF
	E_CIP_Usage.eLine_Color:;
			IF TRUE THEN;
				eProcess:=E_CIP_Usage.eLine_Color;
			END_IF

	E_CIP_Usage.eLine_Marinada:;
			IF TRUE THEN;
				eProcess:=E_CIP_Usage.eLine_Marinada;
			END_IF	
			
	E_CIP_Usage.eLocal:;
			IF TRUE THEN;
				eProcess:=E_CIP_Usage.eLocal;
			END_IF	

	E_CIP_Usage.eNotInUse:;
			IF TRUE THEN;
				eProcess:=E_CIP_Usage.eNotInUse;
			END_IF	
			
	E_CIP_Usage.eTank_1:;
			IF TRUE THEN;
				eProcess:=E_CIP_Usage.eTank_1;
			END_IF	
	E_CIP_Usage.eTank_2:;
			IF TRUE THEN;
				eProcess:=E_CIP_Usage.eTank_2;
			END_IF	
	E_CIP_Usage.eTank_3:;
			IF TRUE THEN;
				eProcess:=E_CIP_Usage.eTank_3;
			END_IF	
	E_CIP_Usage.eTank_4:;
			IF TRUE THEN;
				eProcess:=E_CIP_Usage.eTank_4;
			END_IF	
	E_CIP_Usage.eTriBlender_Color:;
			IF TRUE THEN;
				eProcess:=E_CIP_Usage.eTriBlender_Color;
			END_IF	
	E_CIP_Usage.eTriBlender_Marinada:;
			IF TRUE THEN;
				eProcess:=E_CIP_Usage.eTriBlender_Marinada;
			END_IF	

END_CASE
*)
END_ACTION

ACTION _aReady_exit:
bRun:=TRUE;
bDone:=FALSE;
END_ACTION

ACTION act_GetReference:
m_Set_SFCFlags_Reference();
//refElement REF= fbElement[eElementID];
//refState_Long REF= fbElement[eElementID].eState_Long;

stPis_Client_Source			REF= g_Piston.stPis[valClient_Source];
stPis_Client_Return			REF= g_Piston.stPis[valClient_Return];
stPis_S_Marinade_Up			REF= g_Piston.stPis[valS_Marinade_Up];
//stPis_S_Marinade_Up_Drain	REF= g_Piston.stPis[valS_Marinade_Up_Drain];
stPis_S_Marinade_Low		REF= g_Piston.stPis[valS_Marinade_Low];
stPis_S_Color_Up			REF= g_Piston.stPis[valS_Color_Up];
//stPis_S_Color_Up_Drain		REF= g_Piston.stPis[valS_Color_Up_Drain];
stPis_S_Color_Low			REF= g_Piston.stPis[valS_Color_Low];
//stPis_Tank_1				REF= g_Piston.stPis[valTank_1];
//stPis_Tank_2				REF= g_Piston.stPis[valTank_2];
//stPis_Tank_3				REF= g_Piston.stPis[valTank_3];
//stPis_Tank_4				REF= g_Piston.stPis[valTank_4];
//stPis_S_Marinade_Low_Select	REF= g_Piston.stPis[valS_Marinade_Low_Select];
//stPis_S_Color_Low_Select	REF= g_Piston.stPis[valS_Color_Low_Select];
stPis_Drain					REF= g_Piston.stPis[valDrain];
stPis_Loop				REF= g_Piston.stPis[valLoop];
stPis_S_Future				REF= g_Piston.stPis[valS_Future];
END_ACTION

ACTION act_Oper:
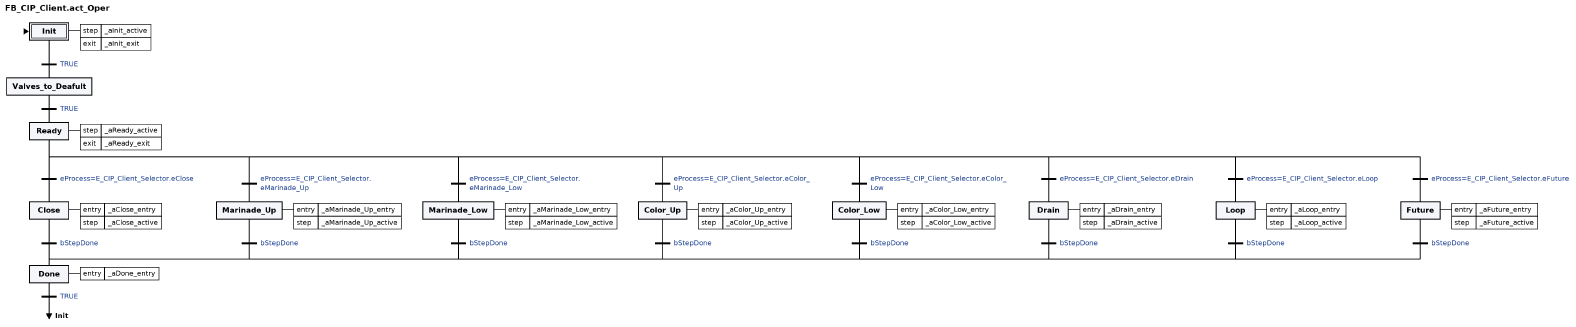
INITIAL_STEP Init:  // min time T#0.5s
    _aInit_active(N);  // step action
    _aInit_exit(P0);  // exit action
END_STEP
TRANSITION FROM Init TO Valves_to_Deafult
    := TRUE;
END_TRANSITION
STEP Valves_to_Deafult:
END_STEP
TRANSITION FROM Valves_to_Deafult TO Ready
    := TRUE;
END_TRANSITION
STEP Ready:
    _aReady_active(N);  // step action
    _aReady_exit(P0);  // exit action
END_STEP
TRANSITION FROM Ready TO Close
    := eProcess=E_CIP_Client_Selector.eClose;
END_TRANSITION
STEP Close:
    _aClose_entry(P1);  // entry action
    _aClose_active(N);  // step action
END_STEP
TRANSITION FROM Close TO Done
    := bStepDone;
END_TRANSITION
TRANSITION FROM Ready TO Marinade_Up
    := eProcess=E_CIP_Client_Selector.eMarinade_Up;
END_TRANSITION
STEP Marinade_Up:
    _aMarinade_Up_entry(P1);  // entry action
    _aMarinade_Up_active(N);  // step action
END_STEP
TRANSITION FROM Marinade_Up TO Done
    := bStepDone;
END_TRANSITION
TRANSITION FROM Ready TO Marinade_Low
    := eProcess=E_CIP_Client_Selector.eMarinade_Low;
END_TRANSITION
STEP Marinade_Low:
    _aMarinade_Low_entry(P1);  // entry action
    _aMarinade_Low_active(N);  // step action
END_STEP
TRANSITION FROM Marinade_Low TO Done
    := bStepDone;
END_TRANSITION
TRANSITION FROM Ready TO Color_Up
    := eProcess=E_CIP_Client_Selector.eColor_Up;
END_TRANSITION
STEP Color_Up:
    _aColor_Up_entry(P1);  // entry action
    _aColor_Up_active(N);  // step action
END_STEP
TRANSITION FROM Color_Up TO Done
    := bStepDone;
END_TRANSITION
TRANSITION FROM Ready TO Color_Low
    := eProcess=E_CIP_Client_Selector.eColor_Low;
END_TRANSITION
STEP Color_Low:
    _aColor_Low_entry(P1);  // entry action
    _aColor_Low_active(N);  // step action
END_STEP
TRANSITION FROM Color_Low TO Done
    := bStepDone;
END_TRANSITION
TRANSITION FROM Ready TO Drain
    := eProcess=E_CIP_Client_Selector.eDrain;
END_TRANSITION
STEP Drain:
    _aDrain_entry(P1);  // entry action
    _aDrain_active(N);  // step action
END_STEP
TRANSITION FROM Drain TO Done
    := bStepDone;
END_TRANSITION
TRANSITION FROM Ready TO Loop
    := eProcess=E_CIP_Client_Selector.eLoop;
END_TRANSITION
STEP Loop:
    _aLoop_entry(P1);  // entry action
    _aLoop_active(N);  // step action
END_STEP
TRANSITION FROM Loop TO Done
    := bStepDone;
END_TRANSITION
TRANSITION FROM Ready TO Future
    := eProcess=E_CIP_Client_Selector.eFuture;
END_TRANSITION
STEP Future:
    _aFuture_entry(P1);  // entry action
    _aFuture_active(N);  // step action
END_STEP
TRANSITION FROM Future TO Done
    := bStepDone;
END_TRANSITION
STEP Done:  // min time T#0.2s
    _aDone_entry(P1);  // entry action
END_STEP
TRANSITION FROM Done TO Init
    := TRUE;
END_TRANSITION
// branch label Branch2_act_Oper
END_ACTION

ACTION act_Status:
IF bReady AND bDone OR TRUE THEN;
	IF TRUE 
	AND fbPis.m_CheckByRecipe(stPis:=stPis_Client_Source, 		req:=E_Piston_Recipe_State.Release)
	AND fbPis.m_CheckByRecipe(stPis:=stPis_Client_Return, 		req:=E_Piston_Recipe_State.Release)
	AND fbPis.m_CheckByRecipe(stPis:=stPis_S_Marinade_Up, 		req:=E_Piston_Recipe_State.Release)
	AND fbPis.m_CheckByRecipe(stPis:=stPis_S_Marinade_Low, 		req:=E_Piston_Recipe_State.Release)
	AND fbPis.m_CheckByRecipe(stPis:=stPis_S_Color_Up, 			req:=E_Piston_Recipe_State.Release)
	AND fbPis.m_CheckByRecipe(stPis:=stPis_S_Color_Low, 		req:=E_Piston_Recipe_State.Release)
	AND fbPis.m_CheckByRecipe(stPis:=stPis_Drain, 				req:=E_Piston_Recipe_State.Release)
	AND fbPis.m_CheckByRecipe(stPis:=stPis_Loop, 				req:=E_Piston_Recipe_State.Release)
	AND fbPis.m_CheckByRecipe(stPis:=stPis_S_Future, 			req:=E_Piston_Recipe_State.Release)
	THEN;
		eStatus:=E_CIP_Client_Selector.eClose;
	ELSIF TRUE
	AND fbPis.m_CheckByRecipe(stPis:=stPis_Client_Source, 		req:=E_Piston_Recipe_State.Act)
	AND fbPis.m_CheckByRecipe(stPis:=stPis_Client_Return, 		req:=E_Piston_Recipe_State.Act)
	AND fbPis.m_CheckByRecipe(stPis:=stPis_S_Marinade_Up, 		req:=E_Piston_Recipe_State.Act)
	AND fbPis.m_CheckByRecipe(stPis:=stPis_S_Marinade_Low, 		req:=E_Piston_Recipe_State.Release)
	AND fbPis.m_CheckByRecipe(stPis:=stPis_S_Color_Up, 			req:=E_Piston_Recipe_State.Release)
	AND fbPis.m_CheckByRecipe(stPis:=stPis_S_Color_Low, 		req:=E_Piston_Recipe_State.Release)
	AND fbPis.m_CheckByRecipe(stPis:=stPis_Drain, 				req:=E_Piston_Recipe_State.Release)
	AND fbPis.m_CheckByRecipe(stPis:=stPis_Loop, 				req:=E_Piston_Recipe_State.Release)
	AND fbPis.m_CheckByRecipe(stPis:=stPis_S_Future, 			req:=E_Piston_Recipe_State.Release)
	THEN;
		eStatus:=E_CIP_Client_Selector.eMarinade_Up;
	ELSIF TRUE 
	AND fbPis.m_CheckByRecipe(stPis:=stPis_Client_Source, 		req:=E_Piston_Recipe_State.Act)
	AND fbPis.m_CheckByRecipe(stPis:=stPis_Client_Return, 		req:=E_Piston_Recipe_State.Act)
	AND fbPis.m_CheckByRecipe(stPis:=stPis_S_Marinade_Up, 		req:=E_Piston_Recipe_State.Release)
	AND fbPis.m_CheckByRecipe(stPis:=stPis_S_Marinade_Low, 		req:=E_Piston_Recipe_State.Act)
	AND fbPis.m_CheckByRecipe(stPis:=stPis_S_Color_Up, 			req:=E_Piston_Recipe_State.Release)
	AND fbPis.m_CheckByRecipe(stPis:=stPis_S_Color_Low, 		req:=E_Piston_Recipe_State.Release)
	AND fbPis.m_CheckByRecipe(stPis:=stPis_Drain, 				req:=E_Piston_Recipe_State.Release)
	AND fbPis.m_CheckByRecipe(stPis:=stPis_Loop, 				req:=E_Piston_Recipe_State.Release)
	AND fbPis.m_CheckByRecipe(stPis:=stPis_S_Future, 			req:=E_Piston_Recipe_State.Release)
	THEN;
		eStatus:=E_CIP_Client_Selector.eMarinade_Low;
	ELSIF TRUE 
	AND fbPis.m_CheckByRecipe(stPis:=stPis_Client_Source, 		req:=E_Piston_Recipe_State.Act)
	AND fbPis.m_CheckByRecipe(stPis:=stPis_Client_Return, 		req:=E_Piston_Recipe_State.Act)
	AND fbPis.m_CheckByRecipe(stPis:=stPis_S_Marinade_Up, 		req:=E_Piston_Recipe_State.Release)
	AND fbPis.m_CheckByRecipe(stPis:=stPis_S_Marinade_Low, 		req:=E_Piston_Recipe_State.Release)
	AND fbPis.m_CheckByRecipe(stPis:=stPis_S_Color_Up, 			req:=E_Piston_Recipe_State.Act)
	AND fbPis.m_CheckByRecipe(stPis:=stPis_S_Color_Low, 		req:=E_Piston_Recipe_State.Release)
	AND fbPis.m_CheckByRecipe(stPis:=stPis_Drain, 				req:=E_Piston_Recipe_State.Release)
	AND fbPis.m_CheckByRecipe(stPis:=stPis_Loop, 				req:=E_Piston_Recipe_State.Release)
	AND fbPis.m_CheckByRecipe(stPis:=stPis_S_Future, 			req:=E_Piston_Recipe_State.Release)
	THEN;
		eStatus:=E_CIP_Client_Selector.eColor_Up;
	ELSIF TRUE 
	AND fbPis.m_CheckByRecipe(stPis:=stPis_Client_Source, 		req:=E_Piston_Recipe_State.Act)
	AND fbPis.m_CheckByRecipe(stPis:=stPis_Client_Return, 		req:=E_Piston_Recipe_State.Act)
	AND fbPis.m_CheckByRecipe(stPis:=stPis_S_Marinade_Up, 		req:=E_Piston_Recipe_State.Release)
	AND fbPis.m_CheckByRecipe(stPis:=stPis_S_Marinade_Low, 		req:=E_Piston_Recipe_State.Release)
	AND fbPis.m_CheckByRecipe(stPis:=stPis_S_Color_Up, 			req:=E_Piston_Recipe_State.Release)
	AND fbPis.m_CheckByRecipe(stPis:=stPis_S_Color_Low, 		req:=E_Piston_Recipe_State.Act)
	AND fbPis.m_CheckByRecipe(stPis:=stPis_Drain, 				req:=E_Piston_Recipe_State.Release)
	AND fbPis.m_CheckByRecipe(stPis:=stPis_Loop, 				req:=E_Piston_Recipe_State.Release)
	AND fbPis.m_CheckByRecipe(stPis:=stPis_S_Future, 			req:=E_Piston_Recipe_State.Release)
	THEN;
		eStatus:=E_CIP_Client_Selector.eColor_Low;
	ELSIF TRUE 
	AND fbPis.m_CheckByRecipe(stPis:=stPis_Client_Source, 		req:=E_Piston_Recipe_State.Release)
	AND fbPis.m_CheckByRecipe(stPis:=stPis_Client_Return, 		req:=E_Piston_Recipe_State.Release)
	AND fbPis.m_CheckByRecipe(stPis:=stPis_S_Marinade_Up, 		req:=E_Piston_Recipe_State.Release)
	AND fbPis.m_CheckByRecipe(stPis:=stPis_S_Marinade_Low, 		req:=E_Piston_Recipe_State.Release)
	AND fbPis.m_CheckByRecipe(stPis:=stPis_S_Color_Up, 			req:=E_Piston_Recipe_State.Release)
	AND fbPis.m_CheckByRecipe(stPis:=stPis_S_Color_Low, 		req:=E_Piston_Recipe_State.Release)
	AND fbPis.m_CheckByRecipe(stPis:=stPis_Drain, 				req:=E_Piston_Recipe_State.Act)
	AND fbPis.m_CheckByRecipe(stPis:=stPis_Loop, 				req:=E_Piston_Recipe_State.Release)
	AND fbPis.m_CheckByRecipe(stPis:=stPis_S_Future, 			req:=E_Piston_Recipe_State.Release)
	THEN;
		eStatus:=E_CIP_Client_Selector.eDrain;
	ELSIF TRUE 
	AND fbPis.m_CheckByRecipe(stPis:=stPis_Client_Source, 		req:=E_Piston_Recipe_State.Act)
	AND fbPis.m_CheckByRecipe(stPis:=stPis_Client_Return, 		req:=E_Piston_Recipe_State.Act)
	AND fbPis.m_CheckByRecipe(stPis:=stPis_S_Marinade_Up, 		req:=E_Piston_Recipe_State.Release)
	AND fbPis.m_CheckByRecipe(stPis:=stPis_S_Marinade_Low, 		req:=E_Piston_Recipe_State.Release)
	AND fbPis.m_CheckByRecipe(stPis:=stPis_S_Color_Up, 			req:=E_Piston_Recipe_State.Release)
	AND fbPis.m_CheckByRecipe(stPis:=stPis_S_Color_Low, 		req:=E_Piston_Recipe_State.Release)
	AND fbPis.m_CheckByRecipe(stPis:=stPis_Drain, 				req:=E_Piston_Recipe_State.Act)
	AND fbPis.m_CheckByRecipe(stPis:=stPis_Loop, 				req:=E_Piston_Recipe_State.Act)
	AND fbPis.m_CheckByRecipe(stPis:=stPis_S_Future, 			req:=E_Piston_Recipe_State.Release)
	THEN;
		eStatus:=E_CIP_Client_Selector.eLoop;
	ELSIF TRUE 
	AND fbPis.m_CheckByRecipe(stPis:=stPis_Client_Source, 		req:=E_Piston_Recipe_State.Act)
	AND fbPis.m_CheckByRecipe(stPis:=stPis_Client_Return, 		req:=E_Piston_Recipe_State.Act)
	AND fbPis.m_CheckByRecipe(stPis:=stPis_S_Marinade_Up, 		req:=E_Piston_Recipe_State.Release)
	AND fbPis.m_CheckByRecipe(stPis:=stPis_S_Marinade_Low, 		req:=E_Piston_Recipe_State.Release)
	AND fbPis.m_CheckByRecipe(stPis:=stPis_S_Color_Up, 			req:=E_Piston_Recipe_State.Release)
	AND fbPis.m_CheckByRecipe(stPis:=stPis_S_Color_Low, 		req:=E_Piston_Recipe_State.Release)
	AND fbPis.m_CheckByRecipe(stPis:=stPis_Drain, 				req:=E_Piston_Recipe_State.Release)
	AND fbPis.m_CheckByRecipe(stPis:=stPis_Loop, 				req:=E_Piston_Recipe_State.Release)
	AND fbPis.m_CheckByRecipe(stPis:=stPis_S_Future, 			req:=E_Piston_Recipe_State.Release)
	THEN;
		eStatus:=E_CIP_Client_Selector.eFuture;
	ELSE;
		eStatus:=E_CIP_Client_Selector.eNone;
	END_IF
ELSE;
	eStatus:=E_CIP_Client_Selector.eNone;
END_IF
END_ACTION

METHOD m_CheckStatus : BOOL
VAR_INPUT
	eReqStatus		: E_CIP_Usage;
END_VAR
VAR
	eReqStatusLocal	: E_CIP_Client_Selector;
END_VAR
CASE eReqStatus OF
	E_CIP_Usage.eExternal:;
				eReqStatusLocal	:=E_CIP_Client_Selector.eFuture;
	E_CIP_Usage.eLocal:;
				eReqStatusLocal	:=E_CIP_Client_Selector.eClose;
	E_CIP_Usage.eTank_1,
	E_CIP_Usage.eTank_2:;
				eReqStatusLocal	:=E_CIP_Client_Selector.eMarinade_Up;	
	E_CIP_Usage.eTank_3,
	E_CIP_Usage.eTank_4:;
				eReqStatusLocal	:=E_CIP_Client_Selector.eColor_Up;	
	E_CIP_Usage.eTriBlender_Marinada,
	E_CIP_Usage.eLine_Marinada:;
				eReqStatusLocal	:=E_CIP_Client_Selector.eMarinade_Low;	
	E_CIP_Usage.eTriBlender_Color,
	E_CIP_Usage.eLine_Color:;
				eReqStatusLocal	:=E_CIP_Client_Selector.eColor_Low;	
	
END_CASE

IF eStatus=eReqStatusLocal 
AND eProcess=E_CIP_Client_Selector.eNone
AND eReq=E_CIP_Client_Selector.eNone
AND bReady
AND bDone
AND NOT bRun
THEN;
	m_CheckStatus:=TRUE;
END_IF
END_METHOD

METHOD m_IsFree : BOOL
// In Ready with no request: a command given now will not be lost
IF eProcess=E_CIP_Client_Selector.eNone
AND eReq=E_CIP_Client_Selector.eNone
AND bReady
AND NOT bRun
THEN;
	m_IsFree:=TRUE;
END_IF
END_METHOD

METHOD m_Request_Reset : BOOL
VAR_IN_OUT
	memo: R_TRIG;
END_VAR
memo(CLK:=eReq=0);
IF TRUE 
AND memo.Q
THEN;
	SFCReset:=TRUE;
END_IF
END_METHOD

METHOD m_Run : BOOL
VAR_INPUT
	eReqProc			: E_CIP_Usage;
END_VAR
VAR
	eReqStatusLocal	: E_CIP_Client_Selector;
END_VAR
CASE eReqProc OF
	E_CIP_Usage.eExternal:;
				eReqStatusLocal	:=E_CIP_Client_Selector.eFuture;
	E_CIP_Usage.eLocal:;
				eReqStatusLocal	:=E_CIP_Client_Selector.eClose;
	E_CIP_Usage.eTank_1,
	E_CIP_Usage.eTank_2:;
				eReqStatusLocal	:=E_CIP_Client_Selector.eMarinade_Up;	
	E_CIP_Usage.eTank_3,
	E_CIP_Usage.eTank_4:;
				eReqStatusLocal	:=E_CIP_Client_Selector.eColor_Up;	
	E_CIP_Usage.eTriBlender_Marinada,
	E_CIP_Usage.eLine_Marinada:;
				eReqStatusLocal	:=E_CIP_Client_Selector.eMarinade_Low;	
	E_CIP_Usage.eTriBlender_Color,
	E_CIP_Usage.eLine_Color:;
				eReqStatusLocal	:=E_CIP_Client_Selector.eColor_Low;	
	
END_CASE

IF eProcess=E_CIP_Client_Selector.eNone THEN;
	eProcess:=eReq:=eReqStatusLocal;
	bDone:=FALSE;
	m_Run:=TRUE;
END_IF
END_METHOD

METHOD m_Set_SFCFlags_Reference : BOOL
//Set reference to SFC flags

refSFC.SFCInit REF= SFCInit;
refSFC.SFCReset REF= SFCReset;
refSFC.SFCError REF= SFCError;
refSFC.SFCEnableLimit REF= SFCEnableLimit;
refSFC.SFCErrorStep REF= SFCErrorStep;
refSFC.SFCErrorPOU REF= SFCErrorPOU;
refSFC.SFCQuitError REF= SFCQuitError;
refSFC.SFCPause REF= SFCPause;
refSFC.SFCTrans REF= SFCTrans;
refSFC.SFCCurrentStep REF= SFCCurrentStep;
refSFC.SFCTip REF= SFCTip;
refSFC.SFCTipMode REF= SFCTipMode;

// Cycle handle for SFC
m_SFC_Handle();
END_METHOD

END_FUNCTION_BLOCK

// ---- 03 Project/23 CIP/FB_CIP.TcPOU
FUNCTION_BLOCK FB_CIP EXTENDS FB_SFC_Cycle IMPLEMENTS ITF_FB_SFC_Cycle
VAR_INPUT
	valFillWater_T91	: E_Pis_Name;
	valFillWater_T92	: E_Pis_Name;
	valFillWater_T93	: E_Pis_Name;
	valFillWater_T94	: E_Pis_Name;
	
	lvlTank_T91			: ST_Tank_Level	;
	lvlTank_T92			: ST_Tank_Level	;
	lvlTank_T93			: ST_Tank_Level	;
	lvlTank_T94			: ST_Tank_Level	;
	
	eCIP_Usage			: E_CIP_Usage;
	nLocalRecipe		: INT;			//recipe of the local preparation: temperature, concentration, tank volumes (Vadim 02.11.2026, item 7)

END_VAR
VAR_OUTPUT
END_VAR
VAR
	//bRun: BOOL;
	eRun: E_CIP_Source;

	eMode			: E_CIP_Mode;
	eCIP_Return		: E_CIP_Return;
	eCIP_Source		: E_CIP_Source;
	
	eReq			: ST_CIP_Request;
	eReqBlank		: ST_CIP_Request;
	eReqLocal		: ST_CIP_Request;
	
	ref_lvlTank_Client		: REFERENCE TO ST_Tank_Level	;

	//bStepDone: BOOL;
	
	iPosSelect_HMI: INT;

	rtPosMoveHMI_Up		: R_TRIG;
	rtPosMoveHMI_Down	: R_TRIG;
	rtPosDeleteHMI		: R_TRIG;
	rtPosDeleteAllHMI	: R_TRIG;
	
	eCIP_State		: E_Element_State_Long;	// stage reached by the running CIP
	bClientRef_done				: BOOL;
	eState_Long_Blank			: E_Element_State_Long;
	
	fbPis						: FB_Piston;
	stPis_FillWater_T91			: REFERENCE TO ST_Piston;
	stPis_FillWater_T92			: REFERENCE TO ST_Piston;
	stPis_FillWater_T93			: REFERENCE TO ST_Piston;
	stPis_FillWater_T94			: REFERENCE TO ST_Piston;
	
	rtReqLocalCIP_Full_HMI: R_TRIG;
	rtReqLocalCIP_Detergent_HMI: R_TRIG;
	rtReqCleanEmpty_HMI: R_TRIG;
	rtModeOff: R_TRIG;
	rtModeManual: R_TRIG;
	rtModeAuto: R_TRIG;
	bTemp: BOOL;
		
	//Process Control
	//concentration
	stDetergent					:	REFERENCE TO ST_ProcessControl	;
	pcDetergent					: 	REFERENCE TO FB_ProcessControl	;	//detergent local
	stDisInfectant				:	REFERENCE TO ST_ProcessControl	;
	pcDisInfectant				: 	REFERENCE TO FB_ProcessControl	;	//detergent local
    //temperature
	stHeatExchanger					:	REFERENCE TO ST_ProcessControl	;
	pcHeatExchanger					: 	REFERENCE TO FB_ProcessControl	;	//	
	stTemperature_Deterg			:	REFERENCE TO ST_ProcessControl	;
	pcTemperature_Deterg			: 	REFERENCE TO FB_ProcessControl	;	//detergent Client	
	stTemperature_Dis				:	REFERENCE TO ST_ProcessControl	;
	pcTemperature_Dis				: 	REFERENCE TO FB_ProcessControl	;//disinfectant local/client
	//temperature client return
	stTemp_ClntReturn				:	REFERENCE TO ST_ProcessControl	;//Client return temperature
	pcTemp_ClntReturn				: 	REFERENCE TO FB_ProcessControl	;//Client return temperature
	
	//flow rate
	stFlow1_Rate					:	REFERENCE TO ST_ProcessControl	;//CIP
	pcFlow1_Rate					: 	REFERENCE TO FB_ProcessControl	;//disinfectant local/client
	stFlow2_Rate					:	REFERENCE TO ST_ProcessControl	;//CIP send
	pcFlow2_Rate					: 	REFERENCE TO FB_ProcessControl	;//disinfectant local/client	return 
	stFlow3_Rate					:	REFERENCE TO ST_ProcessControl	;//CIP send
	pcFlow3_Rate					: 	REFERENCE TO FB_ProcessControl	;//disinfectant local/client	return 
	
	
	
	//colar marinade 
	//pressure
	stP1001_Pressure				:	REFERENCE TO ST_ProcessControl	;
	pcP1001_Pressure				: 	REFERENCE TO FB_ProcessControl	;//CIP //Client
(*
	stP3001_Pressure				:	REFERENCE TO ST_ProcessControl	;
	pcP3001_Pressure				: 	REFERENCE TO FB_ProcessControl	;
	
	stP3002_Pressure				:	REFERENCE TO ST_ProcessControl	;
	pcP3002_Pressure				: 	REFERENCE TO FB_ProcessControl	;	
	
	stP4001_Pressure				:	REFERENCE TO ST_ProcessControl	;
	pcP4001_Pressure				: 	REFERENCE TO FB_ProcessControl	;
	
	stP4002_Pressure				:	REFERENCE TO ST_ProcessControl	;
	pcP4002_Pressure				: 	REFERENCE TO FB_ProcessControl	;	
	
	stTriBlender_Flow				:	REFERENCE TO ST_ProcessControl	;
	pcTriBlender_Flow				: 	REFERENCE TO FB_ProcessControl	;	
	
	stColor_TriB_Conc				:	REFERENCE TO ST_ProcessControl	;
	pcColor_TriB_Conc				: 	REFERENCE TO FB_ProcessControl	;	
	
	stColor_Line_Conc				:	REFERENCE TO ST_ProcessControl	;
	pcColor_Line_Conc				: 	REFERENCE TO FB_ProcessControl	;	
*)	
	
		//OldOne to be deleted
		iStepDone: INT;
		fDetergTarget: REAL:=0.7;
		fDetergDeviation: REAL;
		fDetergLowTolerance: LREAL;
		fDetergHighTolerance: LREAL;
	

	
	bCIP_Condition_Failed: BOOL;
	testTemperature: REAL := 26.0;
	tonr_CIP_Condition: TONR;
	bCIP_Condition_Done: BOOL;
	fReqVolumeT93: REAL := 250;
	delta_T91_Volume: REAL;	// DisInfection
	delta_T92_Volume: REAL;	// Detergent
	delta_T93_Volume: REAL;	// Recycle Water
	delta_T94_Volume: REAL;	// Water
	memo_T91_Level_start: REAL;
	memo_T92_Level_start: REAL;
	memo_T93_Level_start: REAL;
	memo_T94_Level_start: REAL;	
	
	nStepHeat	:	INT		;
	
	bTestPID: BOOL;
	st_CIP_Param		:	ST_CIP_Param	;
	hystCIP_SetPoint: FB_Hysteresis_REAL;
	a: REAL := 0.8;
	b: REAL := 1.2;
	i: E_CIP_Usage;
	tMeasureDelayTime: TIME;
	bLoadDefSetPoints: BOOL;


	
	//Additional water valume if the solution concentration is too high
	rDeltaWater_DeterLocal		:	REAL	;
	rDeltaWater_DeterClient		:	REAL	;
	rDeltaWater_DisInfLocal		:	REAL	;
	rDeltaWater_DisInfClient	:	REAL	;

	rDeluteVolume				: REAL;
	rDeluteVolume_max			: REAL:=900;

	//accumulative actual time for desinfection and detergent condition
	nDeter_CondActTime_Lcl		:	INT	;//Actual condition time in seconds, for local client, detergent
	nDeter_CondActTime_Clnt		:	INT	;//Actual condition time in seconds, for client, detergent
	nDisInf_CondActTime_Lcl		:	INT	;//Actual condition time in seconds, for local client, disinfection
	nDisInf_CondActTime_Clnt	:	INT	;//Actual condition time in seconds, for client, disinfection
	
	bDeter_CondActTime_Lcl_Done		:	BOOL	;
	bDeter_CondActTime_Clnt_Done	:	BOOL	;
	bDisInf_CondActTime_Lcl_Done	:	BOOL	;
	bDisInf_CondActTime_Clnt_Done	:	BOOL	;

	fbHysteresisFillT94: FB_Hysteresis_REAL;
	
	//Choose pipe or sprinkler
	bSprinkler			:	BOOL:=FALSE	;
	tConditionTime		:	INT		;
	//tConditionTemper:	REAL	;
	fFlowRate			:	REAL	;
	//rVolume_Collect	:	REAL	;
	//rVolume_Drain		:	REAL	;
	//rVolume_Recycle	:	REAL	;
	
	_temp: REAL;
	_cond: ARRAY[0..9] OF BOOL;
	tonStepConditionTime: TON;
	bClientTypeIs_Tank: BOOL;
	t_ActMeasureTime: TIME;
	
	volume_Requered	: INT;
	volume_Actual	: INT;

	ton_Concentration_Filter: TON;
	bConcentration_correct: BOOL;
	tonTankLowLevel: TON;
	iCheck: INT;
	iConcentrationDeluteCounter: INT;
END_VAR
//upper lower control
VAR
	nClient			:	INT:=1		;
	nNumOfRetries	:	INT:=5		;
	nNumOfPulses	:	INT:=5		;//Number of pulses per valve seat clean
	nStep_Vlv		:	INT:=0		;
	bValveCleanDone	:	BOOL:=FALSE	;
	nI_1_act_valve			:	INT:=1		;
	nI_2_act_pulses			:	INT:=0		;
	nI_3_act_repeats		:	INT:=1		;//number of repeats
	ActvValve		:	E_Pis_Name	;
	bSeatStatus		:	BOOL:=FALSE	;
	sState			:	STRING		;
	tOn				:	TON			;
	tOff			:	TON			;
	
	nMaxValves		:	INT:=6		;
	
	arTestOverflow: ARRAY[0..5] OF REAL;

END_VAR

VAR_IN_OUT
	fbCIP_Source	: FB_CIP_Source	;
	fbCIP_Return	: FB_CIP_Return	;
	fbCIP_Usage		: FB_CIP_Client	;
	
	//fbTarget					: FB_Tank_Target	;
	//fbLineSource				: FB_Line_Source	;
	//fbLineTarget				: FB_Line_Target	;
	//fbTriBlenderSource		: FB_Line_Source	;
	//fbTriBlenderTarget		: FB_Line_Target	;

	//fb_PumpLine				: FB_Pump	;
	//fb_PumpTriBlender			: FB_Pump	;
	
	//Pumps
	fb_PumpCIP				: FB_Pump;
	fb_PumpDetergent		: FB_DosingPump;
	fb_PumpDisinfection		: FB_DosingPump;
	
	//Heat Exchenger	
	fb_HeatExchenger	:	FB_HeatExchanger	;
	

END_VAR

m_Set_SFCFlags_Reference();
act_GetReference();
act_CallProcessControl();
//act_HeatExchng();
act_SprinklerCondition();
//SUPER^();

//Selecting client for CIP parameters: recipe = CLIENT ID of Siemens, 0 = Local (Vadim 02.11.2026)
IF eReq.eClient=E_CIP_Usage.eExternal AND eReq.nClientId>=1 AND eReq.nClientId<=g_Data.cnRecipeMax THEN;
	st_CIP_Param:=g_Data.arr_CIP_Recipe[eReq.nClientId];
ELSE;
	st_CIP_Param:=g_Data.arr_CIP_Recipe[0];
END_IF
IF nLocalRecipe<0 OR nLocalRecipe>g_Data.cnRecipeMax THEN;
	nLocalRecipe:=0;
END_IF
FOR i:=1 TO E_CIP_Usage.eLocal DO
	g_Data.arr_CIP_Param[i].sName:=TO_STRING(i);
END_FOR

act_Oper();
act_ReqBuffer();
mVolumeMeter();
bValveCleanDone := TRUE; // no mix-proof valves at GAD

rtModeOff(CLK:=eMode=E_CIP_Mode.eOff);
IF rtModeOff.Q THEN;
	SFCReset:=TRUE;
END_IF

rtModeManual(CLK:=eMode=E_CIP_Mode.eManual);
IF rtModeManual.Q THEN;
	bTemp:=TRUE;
END_IF

rtModeAuto(CLK:=eMode=E_CIP_Mode.eAuto);
IF rtModeAuto.Q THEN;
	//SFCReset:=TRUE;
END_IF

IF bRun AND bClientRef_done THEN;
	act_Run();
END_IF


t_ActMeasureTime:=m_MeasureTimeToHMI();
mFillWater();
//IF bMoveStep THEN bMoveStep:=FALSE; END_IF
(*
arTestOverflow[0]:=m_OverFlowCorrect(
rTc:=arTestOverflow[1], 
rAv:=arTestOverflow[2], 
rAc:=arTestOverflow[3]);
*)

ACTION _aCIP1_Conn_Sprinkler_active:
//Spray ball route is set by Siemens
bStepDone:=g_Anybus.fbAnybus.stIn.bSprinklerState;
END_ACTION

ACTION _aCIP1_Conn_Sprinkler_entry:
bSprinkler:=TRUE;

tonr_CIP_Condition(ResetTime:=TRUE);
END_ACTION

ACTION _aCIP1_Done_entry:
m_Set_CIP_State(eState:=E_Element_State_Long.eCIP_1_Rinzed);
END_ACTION

ACTION _aCIP2_Conn_Sprinkler_active:
//Spray ball route is set by Siemens
bStepDone:=g_Anybus.fbAnybus.stIn.bSprinklerState;
END_ACTION

ACTION _aCIP2_Conn_Sprinkler_entry:
//bSprinkler:=TRUE;

tonr_CIP_Condition(ResetTime:=TRUE);
END_ACTION

ACTION _aCIP2_Done_entry:
IF eReq.eClient=E_CIP_Usage.eLocal THEN;
	m_Set_CIP_State(eState:=E_Element_State_Long.eCIP_2_Deterged);
ELSE;
	m_Set_CIP_State(eState:=E_Element_State_Long.eCIP_2_Deterged);
END_IF
END_ACTION

ACTION _aCIP2_Flow_Sprincler_active:
fb_PumpCIP.m_Run(RPM:=pcFlow1_Rate.mRun_PID(Set_Point:=fFlowRate, controlManual:=NOT(fb_PumpCIP.modeAuto)));


IF TRUE 
AND pcFlow1_Rate.mRun()
AND pcFlow2_Rate.mRun()
//AND pcPressure.mRun()
THEN;
	tonStepConditionTime.IN:=TRUE;
ELSE;
	tonStepConditionTime.IN:=FALSE;
END_IF

tonStepConditionTime(PT:=T#10S);
IF tonStepConditionTime.Q THEN;
	bStepDone:=TRUE;
ELSE;
	bStepDone:=FALSE;
END_IF
END_ACTION

ACTION _aCIP2_Flow_Sprincler_entry:
tonStepConditionTime(IN:=FALSE);

m_DashState_done(stage:=E_CIP_DashStage_List.e06_CIP2_Client_Detergent_Condition_Pipe);
m_DashState_activate(stage:=E_CIP_DashStage_List.e07_CIP2_Client_Detergent_Condition_Sprinkler);
END_ACTION

ACTION _aCIP2_If_ClientIsTank_active:
IF bClientTypeIs_Tank THEN;
	bStepDone:=TRUE;
	m_DashState_done(stage:=E_CIP_DashStage_List.e07_CIP2_Client_Detergent_Condition_Sprinkler);
ELSE;
	bStepDone:=FALSE;
	m_DashState_done(stage:=E_CIP_DashStage_List.e06_CIP2_Client_Detergent_Condition_Pipe);
END_IF
END_ACTION

ACTION _aCIP4_Conn_Sprinkler_active:
//Spray ball route is set by Siemens
bStepDone:=g_Anybus.fbAnybus.stIn.bSprinklerState;
END_ACTION

ACTION _aCIP4_Conn_Sprinkler_entry:
//bSprinkler:=TRUE;

tonr_CIP_Condition(ResetTime:=TRUE);
END_ACTION

ACTION _aCIP4_Done_entry:
m_Set_CIP_State(eState:=E_Element_State_Long.eCIP_4_Sanitized);
END_ACTION

ACTION _aCIP4_Flow_Sprincler_active:
fb_PumpCIP.m_Run(RPM:=pcFlow1_Rate.mRun_PID(Set_Point:=fFlowRate, controlManual:=NOT(fb_PumpCIP.modeAuto)));


IF TRUE 
AND pcFlow1_Rate.mRun()
AND pcFlow2_Rate.mRun()
//AND pcPressure.mRun()
THEN;
	tonStepConditionTime.IN:=TRUE;
ELSE;
	tonStepConditionTime.IN:=FALSE;
END_IF

tonStepConditionTime(PT:=T#10S);
IF tonStepConditionTime.Q THEN;
	bStepDone:=TRUE;
ELSE;
	bStepDone:=FALSE;
END_IF
END_ACTION

ACTION _aCIP4_Flow_Sprincler_entry:
tonStepConditionTime(IN:=FALSE);
m_DashState_done(stage:=E_CIP_DashStage_List.e15_CIP4_Client_DisInfection_Condition_Pipe);
m_DashState_activate(stage:=E_CIP_DashStage_List.e16_CIP4_Client_DisInfection_Condition_Sprinkler);
END_ACTION

ACTION _aCIP4_If_ClientIsTank_active:
IF bClientTypeIs_Tank THEN;
	bStepDone:=TRUE;
	m_DashState_done(stage:=E_CIP_DashStage_List.e16_CIP4_Client_DisInfection_Condition_Sprinkler);
ELSE;
	bStepDone:=FALSE;
	m_DashState_done(stage:=E_CIP_DashStage_List.e15_CIP4_Client_DisInfection_Condition_Pipe);
END_IF
END_ACTION

ACTION _aCIP35_Collect_active:
bStepDone:=FALSE;
IF eCIP_State=E_Element_State_Long.eCIP_2_Deterged THEN;
	volume_Requered:= REAL_TO_INT(st_CIP_Param.r_Volume_Collect_Detergent);
	volume_Actual:= REAL_TO_INT(delta_T92_Volume);
ELSIF eCIP_State=E_Element_State_Long.eCIP_4_Sanitized THEN;
	volume_Requered:= REAL_TO_INT(st_CIP_Param.r_Volume_Collect_DisInfection);
	volume_Actual:= REAL_TO_INT(delta_T91_Volume);
END_IF

IF volume_Actual >= volume_Requered THEN;
	bStepDone:=TRUE;
END_IF
END_ACTION

ACTION _aCIP35_Collect_entry:
mVolumeReset_All();
END_ACTION

ACTION _aCIP35_Conn_Sprinkler_active:
//Spray ball route is set by Siemens
bStepDone:=g_Anybus.fbAnybus.stIn.bSprinklerState;
END_ACTION

ACTION _aCIP35_Conn_Sprinkler_entry:
bSprinkler:=TRUE;

tonr_CIP_Condition(ResetTime:=TRUE);
END_ACTION

ACTION _aCIP35_Done_entry:


CASE eCIP_State OF
	E_Element_State_Long.eNotClean:;
			//
	E_Element_State_Long.eCIP_1_Rinzed:;
			//
	E_Element_State_Long.eCIP_2_Deterged:;
			m_Set_CIP_State(eState:=E_Element_State_Long.eCIP_3_Deterged_Clean);	
		
	E_Element_State_Long.eCIP_3_Deterged_Clean:;
			//
	E_Element_State_Long.eCIP_4_Sanitized:;
			m_Set_CIP_State(eState:=E_Element_State_Long.eCIP_5_Done);			
	
END_CASE
END_ACTION

ACTION _aCIP35_Drain_active:
bStepDone:=FALSE;

IF eCIP_State=E_Element_State_Long.eCIP_2_Deterged THEN;
	volume_Requered:= REAL_TO_INT(st_CIP_Param.r_Volume_Drain_Detergent);
	volume_Actual:= REAL_TO_INT(-delta_T94_Volume);
ELSIF eCIP_State=E_Element_State_Long.eCIP_4_Sanitized THEN;
	volume_Requered:= REAL_TO_INT(st_CIP_Param.r_Volume_Drain_DisInfection);
	volume_Actual:= REAL_TO_INT(-delta_T94_Volume);
END_IF

IF volume_Actual >= volume_Requered THEN;
	bStepDone:=TRUE;
END_IF
END_ACTION

ACTION _aCIP35_Drain_entry:
fbCIP_Return.m_Run(eReqProc:=E_CIP_Return.eDrain);
mVolumeReset_All();

CASE eCIP_State OF

	E_Element_State_Long.eCIP_2_Deterged:;
			m_DashState_done(stage:=E_CIP_DashStage_List.e08_CIP3_Detergent_Collect);
			m_DashState_activate(stage:=E_CIP_DashStage_List.e09_CIP3_Detergent_Drain);

	E_Element_State_Long.eCIP_4_Sanitized:;
			m_DashState_done(stage:=E_CIP_DashStage_List.e17_CIP5_DisInfection_Collect);
			m_DashState_activate(stage:=E_CIP_DashStage_List.e18_CIP5_DisInfection_Drain);
			
END_CASE
END_ACTION

ACTION _aClient_tank_IsEmpty_active:
bStepDone:=m_ClientTank_IsEmpty();
END_ACTION

ACTION _aClient_Validation_check_active:
//The route to the client is made by Siemens before REQUEST ON
bStepDone:=eRun<>E_CIP_Source.eNone;
END_ACTION

ACTION _aClientReference_IsValid_entry:

END_ACTION

ACTION _aCondition_CIP1_Client_active:
IF NOT bSprinkler THEN
	//pipe
	tConditionTime	:=st_CIP_Param.t_ConditionR_Water;
	fFlowRate		:=st_CIP_Param.r_Flow_Pipe;
	
ELSE
	//sprinkler
	tConditionTime	:=st_CIP_Param.t_ConditionR_Water_Sprinkler;
	fFlowRate		:=st_CIP_Param.r_Flow_Sprinkler;
END_IF

IF Condition_CIP1_Client.t > SECOND_TO_TIME(st_CIP_Param.t_PumpInitRun) THEN;
	fb_PumpCIP.m_Run(RPM:=pcFlow1_Rate.mRun_PID(Set_Point:=fFlowRate,controlManual:=NOT(fb_PumpCIP.modeAuto)));
END_IF


tonr_CIP_Condition(PT:=SECOND_TO_TIME(tConditionTime));
//
IF bSprinkler THEN;
	IF TRUE 
	AND pcFlow1_Rate.mRun(mRun=>_cond[1])
	//AND pcFlow3_Rate.mRun(mRun=>_cond[2])
	THEN;
		tonr_CIP_Condition.IN:=TRUE;
	ELSE;
		tonr_CIP_Condition.IN:=FALSE;
	END_IF
ELSE;
	IF TRUE 
	AND pcFlow1_Rate.mRun(mRun=>_cond[1])
	//AND pcFlow2_Rate.mRun(mRun=>_cond[2])
	THEN;
		tonr_CIP_Condition.IN:=TRUE;
	ELSE;
		tonr_CIP_Condition.IN:=FALSE;
	END_IF	
	
END_IF
//

IF tonr_CIP_Condition.Q THEN
	bCIP_Condition_Done:=TRUE;
ELSE;
	bCIP_Condition_Done:=FALSE;	
END_IF

IF FALSE  
//AND delta_T93_Volume < -st_CIP_Param.r_Volume_Drain_R_Water 
OR lvlTank_T93.rTankLevel < 250
THEN;
	bCIP_Condition_Failed:=TRUE;
END_IF



(*
// Connect return to R_Water
IF TRUE 
AND lvlTank_T93.rTankLevel<450 
AND fbCIP_Return.m_CheckStatus(eReqStatus:=E_CIP_Return.eDrain)
THEN;
	fbCIP_Return.m_Run(eReqProc:=E_CIP_Return.eT93_R_Water);
ELSE;
	
END_IF



// Connect return to Drain

IF TRUE 
AND lvlTank_T93.rTankLevel>500 // The tank is full
AND fbCIP_Return.m_CheckStatus(eReqStatus:=E_CIP_Return.eT93_R_Water)
THEN;
	fbCIP_Return.m_Run(eReqProc:=E_CIP_Return.eDrain);
ELSE;
	
END_IF
*)


(*
IF TRUE 
AND bCIP_Condition_Done
OR bCIP_Condition_Failed
THEN;

ELSE;
	
END_IF

IF TRUE 
AND pcFlow1_Rate.mRun(mRun=>_cond[1])
AND pcFlow2_Rate.mRun(mRun=>_cond[2])
//AND pcPressure.mRun()
THEN;
	//
ELSE;
	bCIP_Condition_Failed:=TRUE;
END_IF
*)
END_ACTION

ACTION _aCondition_CIP1_Client_entry:
//fbCIP_Return.m_Run(eReqProc:=E_CIP_Return.eT93_R_Water);

fb_PumpCIP.m_Run(RPM:=st_CIP_Param.r_CIP_Pump);


bCIP_Condition_Failed:=FALSE;
bCIP_Condition_Done:=FALSE;
mVolumeReset_All();
END_ACTION

ACTION _aCondition_CIP1_Client_exit:
tonr_CIP_Condition(IN:=FALSE);
END_ACTION

ACTION _aCondition_CIP2_Client_active:
fb_PumpCIP.m_Run(RPM:=pcFlow1_Rate.mRun_PID(Set_Point:=fFlowRate, controlManual:=NOT(fb_PumpCIP.modeAuto)));


IF bSprinkler THEN;
	IF TRUE 
	AND pcFlow1_Rate.mRun(mRun=>_cond[1])
	AND pcFlow3_Rate.mRun(mRun=>_cond[2])
	THEN;
		//
	ELSE;
		bCIP_Condition_Failed:=TRUE;
	END_IF
ELSE;
	IF TRUE 
	AND pcFlow1_Rate.mRun(mRun=>_cond[1])
	AND pcFlow2_Rate.mRun(mRun=>_cond[2])
	THEN;
		//
	ELSE;
		bCIP_Condition_Failed:=TRUE;
	END_IF	
END_IF

pcHeatExchanger.mRun_PID(Set_Point:=st_CIP_Param.r_Temper_Detergent, controlManual:=g_Data.stHeatExchanger.bManual ,mRun_PID=>_temp);
tonr_CIP_Condition(PT:=SECOND_TO_TIME(tConditionTime));
IF TRUE 
AND pcHeatExchanger.mRun_With_SP(Set_Point:=st_CIP_Param.r_Temper_Detergent, mRun_With_SP=>_cond[3])
//AND pcTemperature_Deterg.mRun_With_SP(Set_Point:=g_Data.arr_CIP_Recipe[nLocalRecipe].r_Temper_Detergent, mRun_With_SP=>_cond[4])
AND pcTemp_ClntReturn.mRun_With_SP(Set_Point:=st_CIP_Param.r_Temper_Detergent, mRun_With_SP=>_cond[5])
AND pcDetergent.mRun_With_SP(Set_Point:=st_CIP_Param.r_DetergentConcentration, mRun_With_SP=>_cond[6])
AND measure_Deterg_2.x
AND TRUE
THEN;
	tonr_CIP_Condition.IN:=TRUE;
ELSE;
	tonr_CIP_Condition.IN:=FALSE;
END_IF

IF tonr_CIP_Condition.Q 
AND bValveCleanDone
THEN;
	bCIP_Condition_Done:=TRUE;
ELSE;
	bCIP_Condition_Done:=FALSE;
END_IF



ton_Concentration_Filter(PT:=T#30S, IN:=stDetergent.Control_ON AND NOT stDetergent.OverFlow);
IF TRUE 
AND ton_Concentration_Filter.Q	
THEN;
	bConcentration_correct:=TRUE;
ELSE;
	bConcentration_correct:=FALSE;
END_IF

// Reverce function
(*
IF Deterg_Conc_Client_Done.x 
AND NOT pcDetergent.mRun() 
THEN;
	bCIP_Condition_Failed:=TRUE;
END_IF

IF Temperature_2_Done.x 
//AND NOT pcTemperature_Deterg.mRun()
AND NOT pcTemp_ClntReturn.mRun()
THEN;
	bCIP_Condition_Failed:=TRUE;
END_IF
*)
(*
//ton_CIP_Condition(PT:=T#30S);
IF tConditionTime-nDeter_CondActTime_Clnt>0 THEN
	tonr_CIP_Condition(PT:=SECOND_TO_TIME(tConditionTime-nDeter_CondActTime_Clnt));
	bDeter_CondActTime_Clnt_Done:=FALSE;
ELSE
	bDeter_CondActTime_Clnt_Done:=TRUE;
END_IF

IF TRUE 
AND Deterg_Conc_Client_Done.x
AND Temperature_2_Done.x
AND NOT bDeter_CondActTime_Clnt_Done
AND TRUE
THEN;
	tonr_CIP_Condition.IN:=TRUE;
ELSE;
	nDeter_CondActTime_Clnt:=TIME_TO_INT(tonr_CIP_Condition.ET)/1000;
	tonr_CIP_Condition.IN:=FALSE;
END_IF

IF tonr_CIP_Condition.Q
OR bDeter_CondActTime_Clnt_Done THEN;
	bCIP_Condition_Done:=TRUE;
ELSE;
	bCIP_Condition_Done:=FALSE;
END_IF
*)
END_ACTION

ACTION _aCondition_CIP2_Client_exit:
tonr_CIP_Condition(IN:=FALSE);
END_ACTION

ACTION _aCondition_CIP2_Local_active:
fb_PumpCIP.m_Run(RPM:=pcFlow1_Rate.mRun_PID(Set_Point:=g_Data.arr_CIP_Recipe[0].r_Flow_Pipe,controlManual:=NOT(fb_PumpCIP.modeAuto)));

IF TRUE 
AND pcFlow1_Rate.mRun(mRun=>_cond[1])
AND pcFlow2_Rate.mRun(mRun=>_cond[2])
//AND pcPressure.mRun()
THEN;
	//
ELSE;
	bCIP_Condition_Failed:=TRUE;
END_IF

pcHeatExchanger.mRun_PID(Set_Point:=g_Data.arr_CIP_Recipe[nLocalRecipe].r_Temper_Detergent, controlManual:=g_Data.stHeatExchanger.bManual ,mRun_PID=>_temp);
tonr_CIP_Condition(PT:=SECOND_TO_TIME(g_Data.arr_CIP_Recipe[0].t_ConditionDetergent), ResetTime:=FALSE);
IF TRUE 
AND pcHeatExchanger.mRun_With_SP(Set_Point:=g_Data.arr_CIP_Recipe[nLocalRecipe].r_Temper_Detergent, mRun_With_SP=>_cond[3])
AND pcTemperature_Deterg.mRun_With_SP(Set_Point:=g_Data.arr_CIP_Recipe[nLocalRecipe].r_Temper_Detergent, mRun_With_SP=>_cond[4])
AND pcTemp_ClntReturn.mRun_With_SP(Set_Point:=g_Data.arr_CIP_Recipe[nLocalRecipe].r_Temper_Detergent, mRun_With_SP=>_cond[5])
AND pcDetergent.mRun_With_SP(Set_Point:=g_Data.arr_CIP_Recipe[nLocalRecipe].r_DetergentConcentration, mRun_With_SP=>_cond[6])
AND measure_Deterg.x
AND TRUE
THEN;
	tonr_CIP_Condition.IN:=TRUE;
ELSE;
	tonr_CIP_Condition.IN:=FALSE;
END_IF
	
IF tonr_CIP_Condition.Q THEN;
	bCIP_Condition_Done:=TRUE;
ELSE;
	bCIP_Condition_Done:=FALSE;	
END_IF


ton_Concentration_Filter(PT:=T#30S, IN:=stDetergent.Control_ON AND NOT stDetergent.OverFlow);
IF TRUE 
AND ton_Concentration_Filter.Q	
THEN;
	bConcentration_correct:=TRUE;
ELSE;
	bConcentration_correct:=FALSE;
END_IF

// Reverce function

(*
IF Deterg_Conc_Local_Done.x 
AND NOT pcDetergent.mRun()
THEN;
	bCIP_Condition_Failed:=TRUE;
END_IF

IF Temperature_1_Done.x 
AND (NOT pcTemperature_Deterg.mRun()
	OR NOT pcTemp_ClntReturn.mRun())
THEN;
	bCIP_Condition_Failed:=TRUE;
END_IF
*)

(*
//ton_CIP_Condition(PT:=T#30S);
IF (g_Data.arr_CIP_Recipe[0].t_ConditionDetergent-nDeter_CondActTime_Lcl)>0 THEN
	tonr_CIP_Condition(PT:=SECOND_TO_TIME(g_Data.arr_CIP_Recipe[0].t_ConditionDetergent-nDeter_CondActTime_Lcl));
	bDeter_CondActTime_Lcl_Done:=FALSE;
ELSE
	bDeter_CondActTime_Lcl_Done:=TRUE;
END_IF

IF TRUE 
AND Deterg_Conc_Local_Done.x
AND Temperature_1_Done.x
AND NOT bDeter_CondActTime_Lcl_Done
AND TRUE
THEN;
	tonr_CIP_Condition.IN:=TRUE;
ELSE;
	nDeter_CondActTime_Lcl:=TIME_TO_INT(tonr_CIP_Condition.ET)/1000;
	tonr_CIP_Condition.IN:=FALSE;
END_IF
	
IF tonr_CIP_Condition.Q OR bDeter_CondActTime_Lcl_Done THEN;
	bCIP_Condition_Done:=TRUE;
ELSE;
	bCIP_Condition_Done:=FALSE;	
END_IF

*)
END_ACTION

ACTION _aCondition_CIP2_Local_exit:
tonr_CIP_Condition(IN:=FALSE);
END_ACTION

ACTION _aCondition_CIP4_Client_active:
fb_PumpCIP.m_Run(RPM:=pcFlow1_Rate.mRun_PID(Set_Point:=fFlowRate,controlManual:=NOT(fb_PumpCIP.modeAuto)));


IF bSprinkler THEN;
	IF TRUE 
	AND pcFlow1_Rate.mRun(mRun=>_cond[1])
	AND pcFlow3_Rate.mRun(mRun=>_cond[2])
	THEN;
		//
	ELSE;
		bCIP_Condition_Failed:=TRUE;
	END_IF
ELSE;
	IF TRUE 
	AND pcFlow1_Rate.mRun(mRun=>_cond[1])
	AND pcFlow2_Rate.mRun(mRun=>_cond[2])
	THEN;
		//
	ELSE;
		bCIP_Condition_Failed:=TRUE;
	END_IF	
END_IF

pcHeatExchanger.mRun_PID(Set_Point:=st_CIP_Param.r_Temper_DisInfection, controlManual:=g_Data.stHeatExchanger.bManual ,mRun_PID=>_temp);
tonr_CIP_Condition(PT:=SECOND_TO_TIME(tConditionTime));
IF TRUE 
AND pcHeatExchanger.mRun_With_SP(Set_Point:=st_CIP_Param.r_Temper_DisInfection, mRun_With_SP=>_cond[3])
//AND pcTemperature_Dis.mRun_With_SP(Set_Point:=st_CIP_Param.r_Temper_DisInfection, mRun_With_SP=>_cond[4])
AND pcTemp_ClntReturn.mRun_With_SP(Set_Point:=st_CIP_Param.r_Temper_DisInfection, mRun_With_SP=>_cond[5])
AND measure_Dis_2.x
AND TRUE
THEN;
	tonr_CIP_Condition.IN:=TRUE;
ELSE;
	tonr_CIP_Condition.IN:=FALSE;
END_IF

IF NOT bSprinkler THEN;
	IF pcDisInfectant.mRun_With_SP(Set_Point:=st_CIP_Param.r_DisInfectionConcentration, mRun_With_SP=>_cond[6])
	AND tonr_CIP_Condition.IN
	THEN;
		//tonr_CIP_Condition.IN:=TRUE;
	ELSIF bSprinkler THEN;
		tonr_CIP_Condition.IN:=TRUE;
	ELSE;
		tonr_CIP_Condition.IN:=FALSE;
	END_IF	
END_IF	


IF tonr_CIP_Condition.Q 
AND bValveCleanDone
THEN
	bCIP_Condition_Done:=TRUE;
ELSE;
	bCIP_Condition_Done:=FALSE;	
END_IF


ton_Concentration_Filter(PT:=T#30S, IN:=stDisInfectant.Control_ON AND (NOT stDisInfectant.OverFlow) AND (NOT bSprinkler));
IF TRUE 	
AND ton_Concentration_Filter.Q	
THEN;
	bConcentration_correct:=TRUE;
ELSE;
	bConcentration_correct:=FALSE;
END_IF

// Reverce function
(*
IF Disinfct_Conc_Client_Done.x 
AND NOT pcDisInfectant.mRun()
AND NOT pcTemp_ClntReturn.mRun()
THEN;
	bCIP_Condition_Failed:=TRUE;
END_IF

IF Temperature_Dis_2_Done.x 
AND NOT pcTemperature_Dis.mRun()
THEN;
	bCIP_Condition_Failed:=TRUE;
END_IF


//ton_CIP_Condition(PT:=T#30S);
IF tConditionTime-nDisInf_CondActTime_Clnt>0 THEN
	tonr_CIP_Condition(PT:=SECOND_TO_TIME(tConditionTime-nDisInf_CondActTime_Clnt));
	bDisInf_CondActTime_Clnt_Done:=FALSE;
ELSE
	bDisInf_CondActTime_Clnt_Done:=TRUE;
END_IF
IF TRUE 
AND Disinfct_Conc_Client_Done.x
AND Temperature_Dis_2_Done.x
AND NOT bDisInf_CondActTime_Clnt_Done
AND TRUE
THEN;
	tonr_CIP_Condition.IN:=TRUE;
ELSE;
	nDisInf_CondActTime_Clnt:=TIME_TO_INT(tonr_CIP_Condition.ET)/1000;
	tonr_CIP_Condition.IN:=FALSE;
END_IF

IF tonr_CIP_Condition.Q 
OR bDisInf_CondActTime_Clnt_Done 
THEN;
	bCIP_Condition_Done:=TRUE;
ELSE;
	bCIP_Condition_Done:=FALSE;	
END_IF
*)
END_ACTION

ACTION _aCondition_CIP4_Client_exit:
tonr_CIP_Condition(IN:=FALSE);
END_ACTION

ACTION _aCondition_CIP4_Local_active:
fb_PumpCIP.m_Run(RPM:=pcFlow1_Rate.mRun_PID(Set_Point:=g_Data.arr_CIP_Recipe[0].r_Flow_Pipe,controlManual:=NOT(fb_PumpCIP.modeAuto)));

IF TRUE 
AND pcFlow1_Rate.mRun(mRun=>_cond[1])
AND pcFlow2_Rate.mRun(mRun=>_cond[2])
//AND pcPressure.mRun()
THEN;
	//
ELSE;
	bCIP_Condition_Failed:=TRUE;
END_IF

pcHeatExchanger.mRun_PID(Set_Point:=g_Data.arr_CIP_Recipe[nLocalRecipe].r_Temper_DisInfection, controlManual:=g_Data.stHeatExchanger.bManual ,mRun_PID=>_temp);
tonr_CIP_Condition(PT:=SECOND_TO_TIME(g_Data.arr_CIP_Recipe[0].t_ConditionDisInfection));
IF TRUE 
AND pcHeatExchanger.mRun_With_SP(Set_Point:=g_Data.arr_CIP_Recipe[nLocalRecipe].r_Temper_DisInfection, mRun_With_SP=>_cond[3])
AND pcTemperature_Dis.mRun_With_SP(Set_Point:=g_Data.arr_CIP_Recipe[nLocalRecipe].r_Temper_DisInfection, mRun_With_SP=>_cond[4])
AND pcTemp_ClntReturn.mRun_With_SP(Set_Point:=g_Data.arr_CIP_Recipe[nLocalRecipe].r_Temper_DisInfection, mRun_With_SP=>_cond[5])
AND pcDisInfectant.mRun_With_SP(Set_Point:=g_Data.arr_CIP_Recipe[nLocalRecipe].r_DisInfectionConcentration, mRun_With_SP=>_cond[6])	
AND measure_Dis.x
AND TRUE
THEN;
	tonr_CIP_Condition.IN:=TRUE;
ELSE;
	tonr_CIP_Condition.IN:=FALSE;
END_IF

IF tonr_CIP_Condition.Q THEN
	bCIP_Condition_Done:=TRUE;
ELSE;
	bCIP_Condition_Done:=FALSE;	
END_IF


ton_Concentration_Filter(PT:=T#30S, IN:=stDisInfectant.Control_ON AND NOT stDisInfectant.OverFlow);
IF TRUE 
AND ton_Concentration_Filter.Q	
THEN;
 bConcentration_correct:=TRUE;
ELSE;
 bConcentration_correct:=FALSE;
END_IF

// Reverce function
(*
IF Disinfct_Conc_Local_Done.x 
AND NOT pcDisInfectant.mRun()
THEN;
	bCIP_Condition_Failed:=TRUE;
END_IF

IF Temperature_Dis_1_Done.x 
AND NOT pcTemperature_Dis.mRun()
THEN;
	bCIP_Condition_Failed:=TRUE;
END_IF
*)
(*
//ton_CIP_Condition(PT:=T#30S);
IF g_Data.arr_CIP_Recipe[0].t_ConditionDisInfection-nDisInf_CondActTime_Lcl>0 THEN
	tonr_CIP_Condition(PT:=SECOND_TO_TIME(g_Data.arr_CIP_Recipe[0].t_ConditionDisInfection-nDisInf_CondActTime_Lcl));
	bDisInf_CondActTime_Lcl_Done:=FALSE;
ELSE
	bDisInf_CondActTime_Lcl_Done:=TRUE;
END_IF

IF TRUE 
AND Disinfct_Conc_Local_Done.x
AND Temperature_Dis_1_Done.x
AND NOT bDisInf_CondActTime_Lcl_Done
AND TRUE
THEN;
	tonr_CIP_Condition.IN:=TRUE;
ELSE;
	nDisInf_CondActTime_Lcl:=TIME_TO_INT(tonr_CIP_Condition.ET)/1000;
	tonr_CIP_Condition.IN:=FALSE;
END_IF

IF tonr_CIP_Condition.Q
OR bDisInf_CondActTime_Lcl_Done
THEN
	bCIP_Condition_Done:=TRUE;
ELSE;
	bCIP_Condition_Done:=FALSE;	
END_IF
*)
END_ACTION

ACTION _aCondition_CIP4_Local_exit:
tonr_CIP_Condition(IN:=FALSE);
END_ACTION

ACTION _aCondition_CIP35_Client_active:
IF NOT bSprinkler THEN
	//pipe
	tConditionTime	:=st_CIP_Param.t_ConditionWater;
	fFlowRate		:=st_CIP_Param.r_Flow_Pipe;
	
ELSE
	//sprinkler
	tConditionTime	:=st_CIP_Param.t_ConditionWater_Sprinkler;
	fFlowRate		:=st_CIP_Param.r_Flow_Sprinkler;
END_IF

IF Condition_CIP35_Client.t > SECOND_TO_TIME(st_CIP_Param.t_PumpInitRun) THEN;
	fb_PumpCIP.m_Run(RPM:=pcFlow1_Rate.mRun_PID(Set_Point:=fFlowRate,controlManual:=NOT(fb_PumpCIP.modeAuto)));
END_IF

//Level control

IF FALSE  
OR lvlTank_T94.rTankLevel < 250
THEN;
	bCIP_Condition_Failed:=TRUE;
END_IF


// Connect return to R_Water
IF TRUE 
AND lvlTank_T93.rTankLevel<450 
AND fbCIP_Return.m_CheckStatus(eReqStatus:=E_CIP_Return.eDrain)
THEN;
	fbCIP_Return.m_Run(eReqProc:=E_CIP_Return.eT93_R_Water);
ELSE;
	
END_IF



// Connect return to Drain

IF TRUE 
AND lvlTank_T93.rTankLevel>500 // The tank is full
AND fbCIP_Return.m_CheckStatus(eReqStatus:=E_CIP_Return.eT93_R_Water)
THEN;
	fbCIP_Return.m_Run(eReqProc:=E_CIP_Return.eDrain);
ELSE;
	
END_IF

// Condition
tonr_CIP_Condition(PT:=SECOND_TO_TIME(tConditionTime));
IF bSprinkler THEN;
	IF TRUE 
	AND pcFlow1_Rate.mRun(mRun=>_cond[1])
	//AND pcFlow3_Rate.mRun(mRun=>_cond[2])
	THEN;
		tonr_CIP_Condition.IN:=TRUE;
	ELSE;
		tonr_CIP_Condition.IN:=FALSE;
	END_IF
ELSE;
	IF TRUE 
	AND pcFlow1_Rate.mRun(mRun=>_cond[1])
	//AND pcFlow2_Rate.mRun(mRun=>_cond[2])
	THEN;
		tonr_CIP_Condition.IN:=TRUE;
	ELSE;
		tonr_CIP_Condition.IN:=FALSE;
	END_IF	
	
END_IF

IF tonr_CIP_Condition.Q THEN
	bCIP_Condition_Done:=TRUE;
ELSE;
	bCIP_Condition_Done:=FALSE;	
END_IF

(*
IF TRUE 
AND bCIP_Condition_Done
OR bCIP_Condition_Failed
THEN;

ELSE;
	
END_IF

IF TRUE 
AND pcFlow1_Rate.mRun(mRun=>_cond[1])
AND pcFlow2_Rate.mRun(mRun=>_cond[2])
//AND pcPressure.mRun()
THEN;
	//
ELSE;
	bCIP_Condition_Failed:=TRUE;
END_IF
*)
END_ACTION

ACTION _aCondition_CIP35_Client_entry:
//fbCIP_Return.m_Run(eReqProc:=E_CIP_Return.eT93_R_Water);
bCIP_Condition_Failed:=FALSE;
bCIP_Condition_Done:=FALSE;
mVolumeReset_All();
END_ACTION

ACTION _aCondition_CIP35_Client_exit:
tonr_CIP_Condition(IN:=FALSE);
END_ACTION

ACTION _aConnect_CIP1_Drain_active:
bStepDone:=FALSE;

IF fbCIP_Source.m_CheckStatus(eReqStatus:=E_CIP_Source.eT93_R_Water) 
AND fbCIP_Usage.m_CheckStatus(eReqStatus:=eReq.eClient)
THEN

	bStepDone:=TRUE;
	
END_IF
END_ACTION

ACTION _aConnect_CIP1_Drain_entry:
fbCIP_Source.m_Run(eReqProc:=E_CIP_Source.eT93_R_Water);
fbCIP_Usage.m_Run(eReqProc:=eReq.eClient);



bSprinkler:=FALSE;
END_ACTION

ACTION _aConnect_CIP2_01_active:
bStepDone:=FALSE;
IF fbCIP_Source.m_CheckStatus(eReqStatus:=E_CIP_Source.eT92_Detergent)  
AND fbCIP_Return.m_CheckStatus(eReqStatus:=E_CIP_Return.eT92_Detergent)  
AND fbPis.m_CheckByRecipe(stPis:=stPis_FillWater_T92, req:=E_Piston_Recipe_State.Release) THEN;
	bStepDone:=TRUE;
END_IF
END_ACTION

ACTION _aConnect_CIP2_01_entry:
fbCIP_Source.m_Run(eReqProc:=E_CIP_Source.eT92_Detergent);
fbCIP_Return.m_Run(eReqProc:=E_CIP_Return.eT92_Detergent);
fbPis.m_SetByRecipe(stPis:=stPis_FillWater_T92, req:=E_Piston_Recipe_State.Release);

m_DashState_done(stage:=E_CIP_DashStage_List.e03_CIP2_Local_Detergent_Fill);
m_DashState_activate(stage:=E_CIP_DashStage_List.e04_CIP2_Local_Detergent_Condition);
END_ACTION

ACTION _aConnect_CIP2_02_active:
bStepDone:=FALSE;
IF fbCIP_Return.m_CheckStatus(eReqStatus:=E_CIP_Return.eT92_Detergent)  
//AND fbPis.m_CheckByRecipe(stPis:=stPis_FillWater_T92, req:=E_Piston_Recipe_State.Release) 
THEN;
	bStepDone:=TRUE;
END_IF
END_ACTION

ACTION _aConnect_CIP2_02_entry:
fbCIP_Return.m_Run(eReqProc:=E_CIP_Return.eT92_Detergent);
fbPis.m_SetByRecipe(stPis:=stPis_FillWater_T92, req:=E_Piston_Recipe_State.Release);
//fb_PumpDetergent.m_Auto();
fb_HeatExchenger.m_Auto();

m_DashState_done(stage:=E_CIP_DashStage_List.e05_CIP2_Client_Detergent_Fill);
m_DashState_activate(stage:=E_CIP_DashStage_List.e06_CIP2_Client_Detergent_Condition_Pipe);
END_ACTION

ACTION _aConnect_CIP2_Drain_active:
bStepDone:=FALSE;
IF fbCIP_Usage.m_CheckStatus(eReqStatus:=eReq.eClient)  
AND fbCIP_Return.m_CheckStatus(eReqStatus:=E_CIP_Return.eDrain) 
THEN;

	bStepDone:=TRUE;
	
END_IF
END_ACTION

ACTION _aConnect_CIP2_Drain_entry:
fbCIP_Usage.m_Run(eReqProc:=eReq.eClient);
fbCIP_Return.m_Run(eReqProc:=E_CIP_Return.eDrain);
fb_HeatExchenger.m_Auto();




m_DashState_activate(stage:=E_CIP_DashStage_List.e05_CIP2_Client_Detergent_Fill);
END_ACTION

ACTION _aConnect_CIP4_01_active:
bStepDone:=FALSE;
IF fbCIP_Source.m_CheckStatus(eReqStatus:=E_CIP_Source.eT91_Sanitation)  
AND fbCIP_Return.m_CheckStatus(eReqStatus:=E_CIP_Return.eT91_Sanitation)  
AND fbPis.m_CheckByRecipe(stPis:=stPis_FillWater_T91, req:=E_Piston_Recipe_State.Release) THEN;
	bStepDone:=TRUE;
END_IF
END_ACTION

ACTION _aConnect_CIP4_01_entry:
fbCIP_Source.m_Run(eReqProc:=E_CIP_Source.eT91_Sanitation);
fbCIP_Return.m_Run(eReqProc:=E_CIP_Return.eT91_Sanitation);
fbPis.m_SetByRecipe(stPis:=stPis_FillWater_T91, req:=E_Piston_Recipe_State.Release);
tonr_CIP_Condition(ResetTime:=TRUE);

m_DashState_done(stage:=E_CIP_DashStage_List.e12_CIP4_Local_DisInfection_Fill);
m_DashState_activate(stage:=E_CIP_DashStage_List.e13_CIP4_Local_DisInfection_Condition);
END_ACTION

ACTION _aConnect_CIP4_02_active:
bStepDone:=FALSE;
IF fbCIP_Return.m_CheckStatus(eReqStatus:=E_CIP_Return.eT91_Sanitation)  
//AND fbPis.m_CheckByRecipe(stPis:=stPis_FillWater_T92, req:=E_Piston_Recipe_State.Release) 
THEN;
	bStepDone:=TRUE;
END_IF
END_ACTION

ACTION _aConnect_CIP4_02_entry:
fbCIP_Return.m_Run(eReqProc:=E_CIP_Return.eT91_Sanitation);

m_DashState_done(stage:=E_CIP_DashStage_List.e14_CIP4_Client_DisInfection_Fill);
m_DashState_activate(stage:=E_CIP_DashStage_List.e15_CIP4_Client_DisInfection_Condition_Pipe);
END_ACTION

ACTION _aConnect_CIP4_Drain_active:
bStepDone:=FALSE;
IF fbCIP_Usage.m_CheckStatus(eReqStatus:=eReq.eClient)  
AND fbCIP_Return.m_CheckStatus(eReqStatus:=E_CIP_Return.eDrain) 
THEN;

	bStepDone:=TRUE;
	
END_IF
END_ACTION

ACTION _aConnect_CIP4_Drain_entry:
fbCIP_Usage.m_Run(eReqProc:=eReq.eClient);
fbCIP_Return.m_Run(eReqProc:=E_CIP_Return.eDrain);
fb_HeatExchenger.m_Auto();




m_DashState_activate(stage:=E_CIP_DashStage_List.e14_CIP4_Client_DisInfection_Fill);
END_ACTION

ACTION _aConnect_CIP35_active:
bStepDone:=FALSE;
IF TRUE
AND fbCIP_Source.m_CheckStatus(eReqStatus:=E_CIP_Source.eT94_Water) 
//AND fbCIP_Source.m_CheckStatus(eReqStatus:=E_CIP_Source.eT93_R_Water) 
AND fbCIP_Usage.m_CheckStatus(eReqStatus:=eReq.eClient)  
//AND fbCIP_Return.m_CheckStatus(eReqStatus:=E_CIP_Return.eDrain) 
THEN;

	bStepDone:=TRUE;
	
END_IF

IF bStepDone THEN;
	CASE eCIP_State OF
		E_Element_State_Long.eCIP_2_Deterged:;
				//fbCIP_Return.m_Run(eReqProc:=E_CIP_Return.eT92_Detergent);
				bStepDone:=fbCIP_Return.m_CheckStatus(eReqStatus:=E_CIP_Return.eT92_Detergent);
		E_Element_State_Long.eCIP_4_Sanitized:;
				//fbCIP_Return.m_Run(eReqProc:=E_CIP_Return.eT91_Sanitation);	
				bStepDone:=fbCIP_Return.m_CheckStatus(eReqStatus:=E_CIP_Return.eT91_Sanitation);
	ELSE;
		bStepDone:=FALSE;
	END_CASE	
END_IF
END_ACTION

ACTION _aConnect_CIP35_entry:
fbCIP_Source.m_Run(eReqProc:=E_CIP_Source.eT94_Water);
//Temp solution for T93
//fbCIP_Source.m_Run(eReqProc:=E_CIP_Source.eT93_R_Water);
fbCIP_Usage.m_Run(eReqProc:=eReq.eClient);




CASE eCIP_State OF
	E_Element_State_Long.eCIP_2_Deterged:;
			fbCIP_Return.m_Run(eReqProc:=E_CIP_Return.eT92_Detergent);
		
	E_Element_State_Long.eCIP_4_Sanitized:;
			fbCIP_Return.m_Run(eReqProc:=E_CIP_Return.eT91_Sanitation);				
END_CASE
END_ACTION

ACTION _aConnect_CIP35_R_Water_active:
bStepDone:=FALSE;
IF fbCIP_Return.m_CheckStatus(eReqStatus:=E_CIP_Return.eT93_R_Water)  
THEN;
	bStepDone:=TRUE;
END_IF
END_ACTION

ACTION _aConnect_CIP35_R_Water_entry:
fbCIP_Return.m_Run(eReqProc:=E_CIP_Return.eT93_R_Water);
mVolumeReset_All();

	CASE eCIP_State OF
	
		E_Element_State_Long.eCIP_2_Deterged:;
				m_DashState_done(stage:=E_CIP_DashStage_List.e09_CIP3_Detergent_Drain);
				m_DashState_activate(stage:=E_CIP_DashStage_List.e10_CIP3_Detergent_Clean_Pipe);
	
		E_Element_State_Long.eCIP_4_Sanitized:;
				m_DashState_done(stage:=E_CIP_DashStage_List.e18_CIP5_DisInfection_Drain);
				m_DashState_activate(stage:=E_CIP_DashStage_List.e19_CIP5_DisInfection_Clean_Pipe);
				
	END_CASE
END_ACTION

ACTION _aDeterg_Dose_1_active:

bStepDone:=fb_PumpDetergent.m_RunVolume(Volume:=0.9*(lvlTank_T92.rTankLevel*stDetergent.Deviation*10)); // 10= 1Litr*1000cc/100%
END_ACTION

ACTION _aDeterg_Dose_2_active:

bStepDone:=fb_PumpDetergent.m_RunVolume(Volume:=0.9*(lvlTank_T92.rTankLevel*stDetergent.Deviation*10)); // 10= 1Litr*1000cc/100%
END_ACTION

ACTION _aDeterg_Overflow_1_active:
IF lvlTank_T92.rTankLevel>=rDeluteVolume OR bCIP_Condition_Failed  THEN;	
	bStepDone:=TRUE;
	fbPis.m_SetByRecipe(stPis:=stPis_FillWater_T92, req:=E_Piston_Recipe_State.Release);
ELSE;
	//Fill water
	bStepDone:=FALSE;
	IF NOT arrTanksSens[E_Tank_Name.T92].get_stTankLevel_OverFlow() THEN;
		fbPis.m_SetByRecipe(stPis:=stPis_FillWater_T92, req:=E_Piston_Recipe_State.Act);			
	END_IF	
END_IF
END_ACTION

ACTION _aDeterg_Overflow_1_entry:
rDeltaWater_DeterLocal:=m_OverFlowCorrect(
							rTc:=stDetergent.rSetPoint , //g_Data.arr_CIP_Recipe[nLocalRecipe].r_DetergentConcentration
							rAv:=lvlTank_T92.rTankLevel , 
							rAc:=stDetergent.rValue );

fbPrintErrMessageByID(sModuleDescription:='CIP',sActErrorID:='101x000x101');							
rDeluteVolume:=rDeltaWater_DeterLocal + lvlTank_T92.rTankLevel;

IF rDeluteVolume>rDeluteVolume_max THEN;
	// message
	iConcentrationDeluteCounter:=iConcentrationDeluteCounter+1;
	IF iConcentrationDeluteCounter>3 THEN;
		fbPrintErrMessageByID(sModuleDescription:='eCIP',sActErrorID:='101x000x103');
	ELSE;
		fbPrintErrMessageByID(sModuleDescription:='CIP',sActErrorID:='101x000x102');
	END_IF
	rDeluteVolume:=rDeluteVolume_max;
END_IF
END_ACTION

ACTION _aDeterg_Overflow_2_active:
IF lvlTank_T92.rTankLevel>=rDeluteVolume OR bCIP_Condition_Failed THEN;	
	bStepDone:=TRUE;
	fbPis.m_SetByRecipe(stPis:=stPis_FillWater_T92, req:=E_Piston_Recipe_State.Release);
ELSE;
	//Fill water
	bStepDone:=FALSE;
	IF NOT arrTanksSens[E_Tank_Name.T92].get_stTankLevel_OverFlow() THEN;
		fbPis.m_SetByRecipe(stPis:=stPis_FillWater_T92, req:=E_Piston_Recipe_State.Act);			
	END_IF	
END_IF
END_ACTION

ACTION _aDeterg_Overflow_2_entry:
rDeltaWater_DeterClient:=m_OverFlowCorrect(
							rTc:=stDetergent.rSetPoint , 
							rAv:=lvlTank_T92.rTankLevel , 
							rAc:=stDetergent.rValue );
							
fbPrintErrMessageByID(sModuleDescription:='CIP',sActErrorID:='101x000x101');							
rDeluteVolume:=rDeltaWater_DeterClient + lvlTank_T92.rTankLevel;

IF rDeluteVolume>rDeluteVolume_max THEN;
	// message
	iConcentrationDeluteCounter:=iConcentrationDeluteCounter+1;
	IF iConcentrationDeluteCounter>3 THEN;
		fbPrintErrMessageByID(sModuleDescription:='eCIP',sActErrorID:='101x000x103');
	ELSE;
		fbPrintErrMessageByID(sModuleDescription:='CIP',sActErrorID:='101x000x102');
	END_IF
	rDeluteVolume:=rDeluteVolume_max;
END_IF
END_ACTION

ACTION _aDisconnect_n_Drain_CIP_Client_active:
bStepDone:=FALSE;

IF fbCIP_Source.m_CheckStatus(eReqStatus:=E_CIP_Source.eClose) 
AND fbCIP_Usage.m_CheckStatus(eReqStatus:=E_CIP_Usage.eLocal) 
AND fbCIP_Return.m_CheckStatus(eReqStatus:=E_CIP_Return.eDrain)
THEN

	bStepDone:=TRUE;
	
END_IF
END_ACTION

ACTION _aDisconnect_n_Drain_CIP_Client_entry:
fbCIP_Source.m_Run(eReqProc:=E_CIP_Source.eClose);
fbCIP_Usage.m_Run(eReqProc:=E_CIP_Usage.eLocal);
fbCIP_Return.m_Run(eReqProc:=E_CIP_Return.eDrain);

IF bClientTypeIs_Tank THEN;
	
END_IF
END_ACTION

ACTION _aDisconnect_Old_Client_entry:
eReq:=eReqBlank;
eRun:=E_CIP_Source.eNone;
m_CleanEmpty_Spaces();
END_ACTION

ACTION _aDisinfct_Dose_1_active:

bStepDone:=fb_PumpDisinfection.m_RunVolume(Volume:=0.9*(lvlTank_T91.rTankLevel*stDisInfectant.Deviation*10)); // 10= 1Litr*1000cc/100%
END_ACTION

ACTION _aDisinfct_Dose_2_active:

bStepDone:=fb_PumpDisinfection.m_RunVolume(Volume:=0.9*(lvlTank_T91.rTankLevel*stDisInfectant.Deviation*10)); // 10= 1Litr*1000cc/100%
END_ACTION

ACTION _aDisinfct_Overflow_1_active:
IF lvlTank_T91.rTankLevel>=rDeluteVolume OR bCIP_Condition_Failed  THEN;	
	bStepDone:=TRUE;
	fbPis.m_SetByRecipe(stPis:=stPis_FillWater_T91, req:=E_Piston_Recipe_State.Release);
ELSE;
	//Fill water
	bStepDone:=FALSE;
	IF NOT arrTanksSens[E_Tank_Name.T91].get_stTankLevel_OverFlow() THEN;
		fbPis.m_SetByRecipe(stPis:=stPis_FillWater_T91, req:=E_Piston_Recipe_State.Act);			
	END_IF	
END_IF
END_ACTION

ACTION _aDisinfct_Overflow_1_entry:
rDeltaWater_DisInfLocal:=m_OverFlowCorrect(
								rTc:=stDisInfectant.rSetPoint , //g_Data.arr_CIP_Recipe[nLocalRecipe].r_DisInfectionConcentration
								rAv:=lvlTank_T91.rTankLevel , 
								rAc:=stDisInfectant.rValue );
								
fbPrintErrMessageByID(sModuleDescription:='CIP',sActErrorID:='101x000x111');							
rDeluteVolume:=rDeltaWater_DisInfLocal + lvlTank_T91.rTankLevel;

IF rDeluteVolume>rDeluteVolume_max THEN;
	// message
	iConcentrationDeluteCounter:=iConcentrationDeluteCounter+1;
	IF iConcentrationDeluteCounter>3 THEN;
		fbPrintErrMessageByID(sModuleDescription:='eCIP',sActErrorID:='101x000x113');
	ELSE;
		fbPrintErrMessageByID(sModuleDescription:='CIP',sActErrorID:='101x000x112');
	END_IF
	
	rDeluteVolume:=rDeluteVolume_max;
END_IF
END_ACTION

ACTION _aDisinfct_Overflow_2_active:
IF lvlTank_T91.rTankLevel>=rDeluteVolume OR bCIP_Condition_Failed  THEN;	
	bStepDone:=TRUE;
	fbPis.m_SetByRecipe(stPis:=stPis_FillWater_T91, req:=E_Piston_Recipe_State.Release);
ELSE;
	//Fill water
	bStepDone:=FALSE;
	IF NOT arrTanksSens[E_Tank_Name.T91].get_stTankLevel_OverFlow() THEN;
		fbPis.m_SetByRecipe(stPis:=stPis_FillWater_T91, req:=E_Piston_Recipe_State.Act);			
	END_IF	
END_IF
END_ACTION

ACTION _aDisinfct_Overflow_2_entry:
rDeltaWater_DisInfClient:=m_OverFlowCorrect(
								rTc:=stDisInfectant.rSetPoint , 
								rAv:=lvlTank_T91.rTankLevel , 
								rAc:=stDisInfectant.rValue );
								
fbPrintErrMessageByID(sModuleDescription:='CIP',sActErrorID:='101x000x111');							
rDeluteVolume:=rDeltaWater_DisInfClient + lvlTank_T91.rTankLevel;

IF rDeluteVolume>rDeluteVolume_max THEN;
	// message
	iConcentrationDeluteCounter:=iConcentrationDeluteCounter+1;
	IF iConcentrationDeluteCounter>3 THEN;
		fbPrintErrMessageByID(sModuleDescription:='eCIP',sActErrorID:='101x000x113');
	ELSE;
		fbPrintErrMessageByID(sModuleDescription:='CIP',sActErrorID:='101x000x112');
	END_IF
	
	rDeluteVolume:=rDeluteVolume_max;
END_IF
END_ACTION

ACTION _aDone_entry:
arCIP_RequestBufer[0]:=eReqBlank;
bRun:=FALSE;
END_ACTION

ACTION _aEnd_Check_active:
bStepDone:=FALSE;
IF TRUE 
AND eCIP_State = E_Element_State_Long.eCIP_1_Rinzed
AND eReq.eType = E_CIP_Type.R_Water
AND eReq.eClient<>E_CIP_Usage.eLocal
THEN;
	bStepDone:=TRUE;
	
ELSIF TRUE 
AND eCIP_State = E_Element_State_Long.eCIP_3_Deterged_Clean
AND eReq.eType = E_CIP_Type.Detergent
//AND eReq.eClient=E_CIP_Usage.eLocal
THEN;
	bStepDone:=TRUE;
	
ELSIF TRUE 
AND eCIP_State = E_Element_State_Long.eCIP_5_Done
AND eReq.eType = E_CIP_Type.Full
//AND eReq.eClient<>E_CIP_Usage.eLocal
THEN;
	bStepDone:=TRUE;
	
END_IF
END_ACTION

ACTION _aFill_For_MixProof_CIP2_active:
bStepDone:=TRUE;
END_ACTION

ACTION _aFill_For_MixProof_CIP2_entry:
bSprinkler:=TRUE;
fb_PumpCIP.m_Run(RPM:=st_CIP_Param.r_CIP_Pump);
END_ACTION

ACTION _aFill_For_MixProof_CIP4_active:
bStepDone:=TRUE;
END_ACTION

ACTION _aFill_For_MixProof_CIP4_entry:
bSprinkler:=TRUE;
fb_PumpCIP.m_Run(RPM:=st_CIP_Param.r_CIP_Pump);
END_ACTION

ACTION _aFill_Solution_CIP2_active:
bStepDone:=FALSE;
volume_Requered:= REAL_TO_INT(st_CIP_Param.r_Volume_Solution_Fill);
volume_Actual:= REAL_TO_INT(-delta_T92_Volume);

IF volume_Actual >= volume_Requered THEN;
	bStepDone:=TRUE;
END_IF
END_ACTION

ACTION _aFill_Solution_CIP4_active:
fb_PumpCIP.m_Run(RPM:=st_CIP_Param.r_CIP_Pump);


bStepDone:=FALSE;
volume_Requered:= REAL_TO_INT(st_CIP_Param.r_Volume_Solution_Fill);
volume_Actual:= REAL_TO_INT(-delta_T91_Volume);

IF volume_Actual >= volume_Requered THEN;
	bStepDone:=TRUE;
END_IF
END_ACTION

ACTION _aFill_Solution_CIP4_entry:
mVolumeReset_All();
tonr_CIP_Condition(ResetTime:=TRUE);
END_ACTION

ACTION _aFill_Water_T91_active:
nDisInf_CondActTime_Lcl:=0;
nDisInf_CondActTime_Clnt:=0;
bDisInf_CondActTime_Lcl_Done:=FALSE;
bDisInf_CondActTime_Clnt_Done:=FALSE;

bStepDone:=FALSE;
IF fbCIP_Source.m_CheckStatus(eReqStatus:=E_CIP_Source.eClose) 
AND fbCIP_Usage.m_CheckStatus(eReqStatus:=E_CIP_Usage.eLocal)  
AND fbCIP_Return.m_CheckStatus(eReqStatus:=E_CIP_Return.eDrain)  
//AND fbPis.m_CheckByRecipe(stPis:=stPis_FillWater_T91, req:=E_Piston_Recipe_State.Act) 
THEN;
	//IF eReq.eClient=E_CIP_Usage.eLocal 
	IF lvlTank_T91.e_state=E_Tank_Level.eLL
	AND lvlTank_T91.rTankLevel>g_Data.arr_CIP_Recipe[nLocalRecipe].r_Tank91_Volume//250 // Local requered Level
	THEN;	
		bStepDone:=TRUE;
		fbPis.m_SetByRecipe(stPis:=stPis_FillWater_T91, req:=E_Piston_Recipe_State.Release);
	(*ELSIF lvlTank_T91.e_state=E_Tank_Level.eLL
	AND lvlTank_T91.rTankLevel>g_Data.arr_CIP_Recipe[nLocalRecipe].r_TankLevel_2//300 // Client requered Level
	THEN;
		//Level OK
		bStepDone:=TRUE;
		fbPis.m_SetByRecipe(stPis:=stPis_FillWater_T91, req:=E_Piston_Recipe_State.Release);*)
	ELSE;
		//Fill water
		IF NOT arrTanksSens[E_Tank_Name.T91].get_stTankLevel_OverFlow() THEN;
			fbPis.m_SetByRecipe(stPis:=stPis_FillWater_T91, req:=E_Piston_Recipe_State.Act);			
		END_IF	
	END_IF	
END_IF
END_ACTION

ACTION _aFill_Water_T91_entry:
fbCIP_Source.m_Run(eReqProc:=E_CIP_Source.eClose);
fbCIP_Usage.m_Run(eReqProc:=E_CIP_Usage.eLocal);
fbCIP_Return.m_Run(eReqProc:=E_CIP_Return.eDrain);
bSprinkler:=FALSE;

m_DashState_activate(stage:=E_CIP_DashStage_List.e12_CIP4_Local_DisInfection_Fill);
END_ACTION

ACTION _aFill_Water_T92_active:
//Reset
nDeter_CondActTime_Lcl:=0;
nDeter_CondActTime_Clnt:=0;
bDeter_CondActTime_Lcl_Done:=FALSE;
bDeter_CondActTime_Clnt_Done:=FALSE;

bStepDone:=FALSE;
IF fbCIP_Source.m_CheckStatus(eReqStatus:=E_CIP_Source.eClose) 
AND fbCIP_Usage.m_CheckStatus(eReqStatus:=E_CIP_Usage.eLocal)  
AND fbCIP_Return.m_CheckStatus(eReqStatus:=E_CIP_Return.eDrain)  
THEN;
	//IF eReq.eClient=E_CIP_Usage.eLocal 
	IF lvlTank_T92.e_state=E_Tank_Level.eLL
	AND lvlTank_T92.rTankLevel>st_CIP_Param.r_Tank92_Volume//st_CIP_Param.r_TankLevel_1//st_CIP_Param.r_Deter_92_TankLvl_1 // Local requered Level
	THEN;	
		bStepDone:=TRUE;
		fbPis.m_SetByRecipe(stPis:=stPis_FillWater_T92, req:=E_Piston_Recipe_State.Release);
	(*ELSIF lvlTank_T92.e_state=E_Tank_Level.eLL
	AND lvlTank_T92.rTankLevel>st_CIP_Param.r_TankVolume_1//Client requered Level
	THEN;
		//Level OK
		bStepDone:=TRUE;
		fbPis.m_SetByRecipe(stPis:=stPis_FillWater_T92, req:=E_Piston_Recipe_State.Release);*)
	ELSE;
		//Fill water
		IF NOT arrTanksSens[E_Tank_Name.T92].get_stTankLevel_OverFlow() THEN;
			fbPis.m_SetByRecipe(stPis:=stPis_FillWater_T92, req:=E_Piston_Recipe_State.Act);			
		END_IF	
	END_IF	
END_IF
END_ACTION

ACTION _aFill_Water_T92_entry:
fbCIP_Source.m_Run(eReqProc:=E_CIP_Source.eClose);
fbCIP_Usage.m_Run(eReqProc:=E_CIP_Usage.eLocal);
fbCIP_Return.m_Run(eReqProc:=E_CIP_Return.eDrain);
bSprinkler:=FALSE;
m_DashState_activate(stage:=E_CIP_DashStage_List.e03_CIP2_Local_Detergent_Fill);
END_ACTION

ACTION _aFill_Water_T93_active:
bStepDone:=FALSE;
IF fbCIP_Source.m_CheckStatus(eReqStatus:=E_CIP_Source.eClose) 
AND fbCIP_Usage.m_CheckStatus(eReqStatus:=E_CIP_Usage.eLocal)
AND fbCIP_Return.m_CheckStatus(eReqStatus:=E_CIP_Return.eDrain) 
THEN;
	IF TRUE
	AND (lvlTank_T93.e_state=E_Tank_Level.eLL OR TRUE)
	AND lvlTank_T93.rTankLevel>st_CIP_Param.r_Tank93_Volume//fReqVolumeT93 // Client requered Level
	THEN;
		//Level OK
		bStepDone:=TRUE;
		fbPis.m_SetByRecipe(stPis:=stPis_FillWater_T93, req:=E_Piston_Recipe_State.Release);
	ELSE;
		//Fill water
		IF NOT arrTanksSens[E_Tank_Name.T93].get_stTankLevel_OverFlow() THEN;
			fbPis.m_SetByRecipe(stPis:=stPis_FillWater_T93, req:=E_Piston_Recipe_State.Act);			
		END_IF
	END_IF	
	
END_IF
END_ACTION

ACTION _aFill_Water_T93_Done_active:
bStepDone:=FALSE;
IF fbPis.m_CheckByRecipe(stPis:=stPis_FillWater_T93, req:=E_Piston_Recipe_State.Release) THEN
	bStepDone:=TRUE;
END_IF
END_ACTION

ACTION _aFill_Water_T93_Done_entry:
fbPis.m_SetByRecipe(stPis:=stPis_FillWater_T93, req:=E_Piston_Recipe_State.Release);
END_ACTION

ACTION _aFill_Water_T93_entry:
fbCIP_Source.m_Run(eReqProc:=E_CIP_Source.eClose);
fbCIP_Usage.m_Run(eReqProc:=E_CIP_Usage.eLocal);
fbCIP_Return.m_Run(eReqProc:=E_CIP_Return.eDrain);



m_DashState_activate(stage:=E_CIP_DashStage_List.e01_CIP1_Client_Drain_Product_Rest_Pipe);
(*
arCIP_DashStage_list[E_CIP_DashStage_List.e01_CIP1_Client_Drain_Product_Rest_Pipe]:=E_CIP_DashStage.eCIPStage_Active;
eCIP_DashStage_actual:=E_CIP_DashStage_List.e01_CIP1_Client_Drain_Product_Rest_Pipe;
sCIP_DashStage_actual:=TO_STRING(eCIP_DashStage_actual);
*)
END_ACTION

ACTION _aFill_Water_T94_active:
bStepDone:=FALSE;
IF fbCIP_Source.m_CheckStatus(eReqStatus:=E_CIP_Source.eClose) 
AND fbCIP_Usage.m_CheckStatus(eReqStatus:=E_CIP_Usage.eLocal)  
AND fbCIP_Return.m_CheckStatus(eReqStatus:=E_CIP_Return.eDrain)  
THEN;//need something in case there are error in level sensor, should jump into error step and close all valves

	//IF eReq.eClient=E_CIP_Usage.eLocal 
	IF TRUE 
	AND (lvlTank_T94.e_state=E_Tank_Level.eLL OR TRUE)
	AND lvlTank_T94.rTankLevel>st_CIP_Param.r_Tank94_Volume//st_CIP_Param.r_Water_TankLvl_Lcl_1 // Client requered Level
	THEN;	
		bStepDone:=TRUE;
		fbPis.m_SetByRecipe(stPis:=stPis_FillWater_T94, req:=E_Piston_Recipe_State.Release);
	ELSE;
		//Fill water
		IF NOT arrTanksSens[E_Tank_Name.T94].get_stTankLevel_OverFlow() THEN;
			fbPis.m_SetByRecipe(stPis:=stPis_FillWater_T94, req:=E_Piston_Recipe_State.Act);			
		END_IF	END_IF	

END_IF
END_ACTION

ACTION _aFill_Water_T94_Done_active:
bStepDone:=FALSE;
IF fbPis.m_CheckByRecipe(stPis:=stPis_FillWater_T94, 		req:=E_Piston_Recipe_State.Act) THEN
	bStepDone:=TRUE;
END_IF
bStepDone:=TRUE;
END_ACTION

ACTION _aFill_Water_T94_Done_entry:
fbPis.m_SetByRecipe(stPis:=stPis_FillWater_T94, 			req:=E_Piston_Recipe_State.Release);
END_ACTION

ACTION _aFill_Water_T94_entry:
fbCIP_Source.m_Run(eReqProc:=E_CIP_Source.eClose);
fbCIP_Usage.m_Run(eReqProc:=E_CIP_Usage.eLocal);
fbCIP_Return.m_Run(eReqProc:=E_CIP_Return.eDrain);
fbPis.m_SetByRecipe(stPis:=stPis_FillWater_T94, 			req:=E_Piston_Recipe_State.Act);


CASE eCIP_State OF

	E_Element_State_Long.eCIP_2_Deterged:;
			m_DashState_activate(stage:=E_CIP_DashStage_List.e08_CIP3_Detergent_Collect);

	E_Element_State_Long.eCIP_4_Sanitized:;
			m_DashState_activate(stage:=E_CIP_DashStage_List.e17_CIP5_DisInfection_Collect);
			
END_CASE
END_ACTION

ACTION _aFlow_Volume_Meter_active:
//

IF eReq.eClient=E_CIP_Usage.eLocal THEN;
	//
ELSE;
	
END_IF

(*

eReq.eClient=E_CIP_Usage.eLocal
*)
END_ACTION

ACTION _aGet_Client_active:
//Next CIP stage
bStepDone:=FALSE;
CASE eReq.eType OF
	E_CIP_Type.R_Water:;
		CASE eCIP_State OF
			E_Element_State_Long.eNotClean:;
					eRun:=E_CIP_Source.eT93_R_Water;
		END_CASE

	E_CIP_Type.Detergent:;
		CASE eCIP_State OF
			E_Element_State_Long.eNotClean:;
					eRun:=E_CIP_Source.eT93_R_Water;

			E_Element_State_Long.eCIP_1_Rinzed:;
					eRun:=E_CIP_Source.eT92_Detergent;

			E_Element_State_Long.eCIP_2_Deterged:;
					eRun:=E_CIP_Source.eT94_Water;
		END_CASE

	E_CIP_Type.Full:;
		CASE eCIP_State OF
			E_Element_State_Long.eNotClean:;
					eRun:=E_CIP_Source.eT93_R_Water;

			E_Element_State_Long.eCIP_1_Rinzed:;
					eRun:=E_CIP_Source.eT92_Detergent;

			E_Element_State_Long.eCIP_2_Deterged:;
					eRun:=E_CIP_Source.eT94_Water;

			E_Element_State_Long.eCIP_3_Deterged_Clean:;
					eRun:=E_CIP_Source.eT91_Sanitation;

			E_Element_State_Long.eCIP_4_Sanitized:;
					eRun:=E_CIP_Source.eT94_Water;
		END_CASE

END_CASE
bStepDone:=TRUE;
END_ACTION

ACTION _aGet_Client_exit:
m_DashState_ToString_convertion();
m_DashState_Get_ToBeDone_List();
END_ACTION

ACTION _ainit_active:
SFCReset:=FALSE;
END_ACTION

ACTION _ainit_exit:
bRun:=FALSE;
IF eMode=E_CIP_Mode.eAuto THEN;
	eMode:=E_CIP_Mode.eManual;
END_IF
g_Data.b_CIP_Run:=FALSE;
_aGet_Client_active();
END_ACTION

ACTION _ameasure_Deterg_2_active:

END_ACTION

ACTION _ameasure_Deterg_active:

END_ACTION

ACTION _ameasure_Dis_2_active:

END_ACTION

ACTION _ameasure_Dis_active:

END_ACTION

ACTION _ameasureDelay_CIP2_1_active:
bStepDone:=FALSE;
tMeasureDelayTime:=SECOND_TO_TIME(g_Data.arr_CIP_Recipe[0].t_Measure_Delay);
IF measureDelay_CIP2_1.t > tMeasureDelayTime THEN;
	bStepDone:=TRUE;
END_IF

IF bCIP_Condition_Failed THEN;
	bStepDone:=TRUE;
END_IF
END_ACTION

ACTION _ameasureDelay_CIP2_1_entry:
pcDetergent.mReset();
END_ACTION

ACTION _ameasureDelay_CIP2_2_active:
bStepDone:=FALSE;
tMeasureDelayTime:=SECOND_TO_TIME(st_CIP_Param.t_Measure_Delay);
IF measureDelay_CIP2_2.t > tMeasureDelayTime THEN;
	bStepDone:=TRUE;
END_IF

IF bCIP_Condition_Failed THEN;
	bStepDone:=TRUE;
END_IF
END_ACTION

ACTION _ameasureDelay_CIP2_2_entry:
pcDetergent.mReset();
END_ACTION

ACTION _ameasureDelay_CIP4_1_active:
bStepDone:=FALSE;
tMeasureDelayTime:=SECOND_TO_TIME(g_Data.arr_CIP_Recipe[0].t_Measure_Delay);
IF measureDelay_CIP4_1.t > tMeasureDelayTime THEN;
	bStepDone:=TRUE;
END_IF

IF bCIP_Condition_Failed THEN;
	bStepDone:=TRUE;
END_IF
END_ACTION

ACTION _ameasureDelay_CIP4_1_entry:
pcDisInfectant.mReset();
END_ACTION

ACTION _ameasureDelay_CIP4_2_active:
bStepDone:=FALSE;
tMeasureDelayTime:= SECOND_TO_TIME(st_CIP_Param.t_Measure_Delay);
IF measureDelay_CIP4_2.t > tMeasureDelayTime 
OR bSprinkler
THEN;
	bStepDone:=TRUE;
END_IF

IF bCIP_Condition_Failed THEN;
	bStepDone:=TRUE;
END_IF
END_ACTION

ACTION _ameasureDelay_CIP4_2_entry:
pcDisInfectant.mReset();
END_ACTION

ACTION _aReady_active:
CASE eMode OF
	E_CIP_Mode.eOff:;
		bRun:=FALSE;
		bStepDone:=FALSE;
	E_CIP_Mode.eManual:;
		IF TRUE 
		AND bRun 
		AND arCIP_RequestBufer[0].eClient<>E_CIP_Usage.eNotInUse
		
		THEN;
			bStepDone:=TRUE;
		ELSE;
			bStepDone:=FALSE;
		END_IF	
	E_CIP_Mode.eAuto:;
		IF TRUE 
		//AND bRun 
		AND arCIP_RequestBufer[0].eClient<>E_CIP_Usage.eNotInUse
		
		THEN;
			bRun:=TRUE;
			bStepDone:=TRUE;
		ELSE;
			bStepDone:=FALSE;
		END_IF		
END_CASE
END_ACTION

ACTION _aReady_exit:
eReq:=arCIP_RequestBufer[0];
bClientTypeIs_Tank:=eReq.eClient=E_CIP_Usage.eExternal AND eReq.eClientType=E_Anybus_ClientType.eTank;

